// TwinCAT 3 PLC project PmsStd
// ProgramVersion: 3.1.4024.0
// libraries:
//   Tc3_IotBase, * (Beckhoff Automation GmbH)
//   Tc2_ModbusRTU, * (Beckhoff Automation GmbH)
//   Tc2_ModbusSrv, * (Beckhoff Automation GmbH)
//   Tc2_Standard, * (Beckhoff Automation GmbH)
//   Tc2_SUPS, * (Beckhoff Automation GmbH)
//   Tc2_System, * (Beckhoff Automation GmbH)
//   Tc3_Module, * (Beckhoff Automation GmbH)
//   Tc3_EventLogger, * (Beckhoff Automation GmbH)
//   Tc2_Utilities, * (Beckhoff Automation GmbH)
// project tree:
//   / FastTask.TcTTO, MqttTask.TcTTO, PlcTask.TcTTO, RedundancyTask.TcTTO
//   10_Core/00_Type/ ST_RuleTargetReg.TcDUT, ST_UnitLimitView.TcDUT, ST_BatLimitView.TcDUT, ST_BatLimitOut.TcDUT, ST_GateView.TcDUT, ST_GateOut.TcDUT, ST_SelectCand.TcDUT, ST_SelectView.TcDUT, ST_DistView.TcDUT, E_GridMode.TcDUT, ST_LogSet.TcDUT, E_StartMode.TcDUT, E_BatClose.TcDUT, ST_SeqSet.TcDUT, E_DistBasis.TcDUT, ST_CmdFilterSet.TcDUT, ST_RedSet.TcDUT, E_RedRole.TcDUT, ST_ModeSet.TcDUT, E_SelectMode.TcDUT, ST_GroupSet.TcDUT, ST_ManualPolicy.TcDUT, GVL_REASON.TcGVL, GVL_CORE.TcGVL, ST_UnitReq.TcDUT, ST_BmsCfg.TcDUT, E_PcsAction.TcDUT, E_BatAction.TcDUT, E_ModeAction.TcDUT, ST_ProtCfg.TcDUT, ST_PointTerm.TcDUT, ST_PointCfg.TcDUT, E_GroupState.TcDUT, E_LimitBasis.TcDUT, E_OpMode.TcDUT, E_ProtScope.TcDUT, E_RunState.TcDUT, E_SourceMode.TcDUT, ST_BatState.TcDUT, ST_GroupCfg.TcDUT, ST_GroupView.TcDUT, ST_Limit.TcDUT, ST_LimitOut.TcDUT, ST_MeterState.TcDUT, ST_ModuleReg.TcDUT, ST_PQ.TcDUT, ST_PccMeas.TcDUT, ST_RuleCfg.TcDUT, ST_SourceOutput.TcDUT, ST_SourceReg.TcDUT, E_PcsCmd.TcDUT, E_BatCmd.TcDUT, ST_PcsCmd.TcDUT, ST_BatCmd.TcDUT, ST_PcsReq.TcDUT, ST_BatReq.TcDUT, ST_PcsSeqSet.TcDUT, ST_BatSeqSet.TcDUT, ST_ManualCmdSet.TcDUT, ST_StateModeSet.TcDUT, ST_PcsCmdMode.TcDUT, ST_BatCmdMode.TcDUT, ST_UnitCfg.TcDUT, ST_UnitState.TcDUT, ST_Val.TcDUT, ST_OutputCfg.TcDUT, ST_ProtReq.TcDUT, ST_ProtView.TcDUT, E_CtrlModeRefuse.TcDUT, E_CtrlModeStep.TcDUT, ST_CtrlModeOut.TcDUT, ST_CtrlModeSet.TcDUT, ST_LocalTime.TcDUT, ST_CtrlModeView.TcDUT, E_PccShare.TcDUT, ST_UnitView.TcDUT
//   10_Core/01_Interface/ I_UnitLimitRule.TcIO, I_BatLimitRule.TcIO, I_Gate.TcIO, I_SelectPolicy.TcIO, I_DistPolicy.TcIO, I_AuxDevice.TcIO, I_OutputRule.TcIO, I_Bms.TcIO, I_CommandSource.TcIO, I_Compensator.TcIO, I_LimitRule.TcIO, I_Meter.TcIO, I_Module.TcIO, I_Pcs.TcIO, I_ReqDevice.TcIO, I_ProtResponse.TcIO, I_ProtectionRule.TcIO, I_StartPermit.TcIO, I_ControlMode.TcIO
//   10_Core/40_Arbitration/ FB_GateAuto.TcPOU, FB_GateManual.TcPOU, FB_SelectStd.TcPOU, F_RangeAnd.TcPOU, FB_PermitEval.TcPOU, FB_OutputReady.TcPOU, E_ModeSwitch.TcDUT, E_ModeStep.TcDUT, E_CmdRefuse.TcDUT, F_CmdOk.TcPOU, FB_ModeSwitch.TcPOU, FB_Gate.TcPOU, E_UnitRole.TcDUT, ST_Pick.TcDUT, ST_Range.TcDUT, ST_Clamp.TcDUT, ST_ShapeDiag.TcDUT, F_LimitKeepZero.TcPOU, F_RangeOpen.TcPOU, F_RangeAdd.TcPOU, F_RangeClamp.TcPOU, F_MakeLimit.TcPOU, F_SourceAllowed.TcPOU, F_StateRank.TcPOU, F_Better.TcPOU, FB_StateArbiter.TcPOU, FB_Select.TcPOU, FB_LimitEval.TcPOU, FB_ShapePath.TcPOU, F_PcsCmdAllowed.TcPOU, F_BatCmdAllowed.TcPOU
//   10_Core/50_Distribution/ FB_DistStd.TcPOU, E_UnitLimitBy.TcDUT, ST_UnitDiag.TcDUT, ST_DistDiag.TcDUT, ST_DistPathDiag.TcDUT, ST_BatDistDiag.TcDUT, FB_Distributor.TcPOU
//   10_Core/20_Protection/ ST_UnitEnvelope.TcDUT, ST_BatEnvelope.TcDUT, ST_GroupEnvelope.TcDUT, FB_EquipmentLimits.TcPOU, ST_BmsProt.TcDUT, ST_BmsAvail.TcDUT, ST_BatGroupState.TcDUT, FB_BatGroup.TcPOU, ST_UnitProt.TcDUT, ST_UnitAvail.TcDUT, F_PcsRank.TcPOU, F_BatRank.TcPOU, FB_Protection.TcPOU, FB_UnitAvail.TcPOU
//   20_Module/Common/ ST_SocLimitSet.TcDUT, ST_RuleBitSet.TcDUT, ST_RuleValueSet.TcDUT, FB_BreakerCtrl.TcPOU, ST_UnitLimitSet.TcDUT, ST_UnitLimitItem.TcDUT, FB_UnitLimit.TcPOU, ST_BreakerSet.TcDUT, F_SocDerate.TcPOU, FB_SocLimit.TcPOU, FB_AuxIo.TcPOU, FB_RuleBit.TcPOU, FB_RuleValue.TcPOU, F_SocLimitSetErr.TcPOU, FB_LocalClock.TcPOU, F_WordsToReal.TcPOU, ST_TempHumState.TcDUT
//   90_Project/ ST_ModuleSet.TcDUT, GVL_TEST.TcGVL, GVL_MQTT.TcGVL, GVL_PARAM.TcGVL, GVL_PERSIST.TcGVL, GVL_SITE.TcGVL, MAIN.TcPOU, GVL_IF.TcGVL, PRG_Mqtt.TcPOU, PRG_Fast.TcPOU, PRG_Redundancy.TcPOU
//   10_Core/60_Dispatch/ FB_GroupState.TcPOU, FB_BatRequest.TcPOU, E_UnitSeq.TcDUT, E_SeqRefuse.TcDUT, F_CmdReached.TcPOU, FB_UnitSeq.TcPOU, FB_BmsSeq.TcPOU, FB_Sequencer.TcPOU, FB_Dispatcher.TcPOU, FB_AuxOutput.TcPOU
//   10_Core/70_Diag/ FB_SettingGuard.TcPOU, FB_ModuleList.TcPOU, E_DiagStage.TcDUT, ST_OutputDiag.TcDUT, E_TraceStep.TcDUT, ST_TraceStep.TcDUT, ST_PTrace.TcDUT, F_TxtPcsAction.TcPOU, F_TxtBatAction.TcPOU, F_TxtSeq.TcPOU, F_TxtRefuse.TcPOU, F_TxtLimitBy.TcPOU, F_TxtStage.TcPOU, F_TxtOpMode.TcPOU, F_TxtCoreReason.TcPOU, F_TxtNum.TcPOU, FB_LogAlarm.TcPOU, FB_LogMsg.TcPOU, FB_OutputDiag.TcPOU, FB_AliveRecorder.TcPOU, FB_EventLog.TcPOU, FB_ConfigCheck.TcPOU, F_TxtPcsCmd.TcPOU, F_TxtBatCmd.TcPOU
//   10_Core/80_Report/ FB_Report.TcPOU
//   10_Core/02_Util/ F_ModeApplies.TcPOU, F_RampStep.TcPOU, FB_Lpf.TcPOU, FB_PersistSave.TcPOU, FB_ReadTimer.TcPOU, F_CycleSec.TcPOU, F_IsStopped.TcPOU, F_IsLocal.TcPOU, F_TimeHhmm.TcPOU, F_RealChanged.TcPOU, F_RealOk.TcPOU, F_RealToDint.TcPOU, F_HhmmOk.TcPOU, F_InHhmmWindow.TcPOU, F_MinutesTo.TcPOU, F_IsFinite.TcPOU
//   10_Core/30_Request/ FB_GroupView.TcPOU, FB_SourceHub.TcPOU, FB_CtrlModeMgr.TcPOU, FB_UnitView.TcPOU
//   20_Module/Standard/ FB_ProtRespStd.TcPOU, FB_ProtPcsFault.TcPOU, FB_ProtPcsComm.TcPOU, FB_ProtBmsFault.TcPOU, FB_ProtBmsComm.TcPOU, FB_ProtPccInvalid.TcPOU
//   10_Core/10_Snapshot/ ST_VirtualSet.TcDUT, FB_Snapshot.TcPOU, FB_Measure.TcPOU
//   10_Core/03_Base/ FB_DeviceBase.TcPOU, FB_ModuleBase.TcPOU, FB_SourceBase.TcPOU, FB_CtrlModeBase.TcPOU
//   20_Module/Mqtt/ FB_MqttPublish.TcPOU, FB_MqttSubscribe.TcPOU, F_MqttDistribute.TcPOU, PRG_PublishDeviceNo.TcPOU, ST_MqttCommand_Rx.TcDUT, ST_MqttCommandHeader.TcDUT, ST_MqttHeader.TcDUT, ST_MqttPubEntry.TcDUT, ST_MqttSubEntry.TcDUT, ST_IfEmsCmd.TcDUT, FB_EmsCommand.TcPOU, FB_SrcEms.TcPOU, FB_MqttMain.TcPOU, ST_MqttBroker.TcDUT, ST_MqttSet.TcDUT, ST_IfReport.TcDUT, F_MqttTimeText.TcPOU, FB_EmsConfigApply.TcPOU, FB_BrokerWatch.TcPOU, E_MqttBroker.TcDUT, ST_BrokerWatchSet.TcDUT, ST_IfEmsCfg.TcDUT, ST_IfEmsCfgEcho.TcDUT, ST_IfUpsConfigRx.TcDUT, FB_EmsCmdGate.TcPOU
//   20_Module/Mqtt/Publish/ ST_AirConditionerPublish_V1.TcDUT, ST_BatPublish_V1.TcDUT, ST_EssPublish_V1.TcDUT, ST_PcsPublish_V1.TcDUT, ST_PmsPublish_V1.TcDUT, ST_PvPublish_V1.TcDUT, ST_RackPublish_V1.TcDUT, ST_TempPublish_V1.TcDUT, ST_AirConditionerPublishData.TcDUT, ST_BatPublishData.TcDUT, ST_EssPublishData.TcDUT, ST_PcsPublishData.TcDUT, ST_PmsPublishData.TcDUT, ST_PvPublishData.TcDUT, ST_RackPublishData.TcDUT, ST_TempPublishData.TcDUT, ST_UpsPublish_V1.TcDUT, ST_ModulePublish_V1.TcDUT, ST_UpsPublishData.TcDUT, ST_ModulePublishData.TcDUT, ST_ImdPublish_V1.TcDUT, ST_ImdPublishData.TcDUT, ST_FirePublish_V1.TcDUT, ST_FirePublishData.TcDUT
//   20_Module/Mqtt/Config/ ST_BatConfig_Rx.TcDUT, ST_CommonConfig_REAL.TcDUT, ST_CommonConfig_UDINT.TcDUT, ST_PcsConfig_Rx.TcDUT, ST_ProtectionConfig_Rx.TcDUT, ST_BatConfigWirePacket.TcDUT, ST_PcsConfigWirePacket.TcDUT, ST_ProtectionConfigWirePacket.TcDUT, ST_UpsConfig_Rx.TcDUT, ST_UpsConfigWirePacket.TcDUT, ST_ScheduleWork_V1.TcDUT, ST_ScheduleHoliday_V1.TcDUT, ST_ScheduleDaily_V1.TcDUT, ST_ScheduleWeekly_V1.TcDUT
//   20_Module/Virtual/ PRG_MqttTestData.TcPOU, FB_BmsSim.TcPOU, FB_MeterSim.TcPOU, FB_PcsSim.TcPOU, FB_SrcTest.TcPOU, PRG_SimLink.TcPOU
//   20_Module/Mqtt/Logger/ FB_MqttLoggerListener.TcPOU, F_Utf8ToWstring.TcPOU, ST_LoggerHeader.TcDUT, ST_LoggerPublish_V1.TcDUT, ST_LoggerSlot.TcDUT
//   20_Module/Report/ FB_RptEsolutionBat.TcPOU, FB_RptSebangUps.TcPOU, FB_RptPlaspoPcs.TcPOU, FB_RptLsImd1000.TcPOU, FB_RptTempHum.TcPOU
//   20_Module/ControlMode/ ST_CmConstPowerSet.TcDUT, FB_CmConstPower.TcPOU, FB_CmStdSchedule.TcPOU, ST_CmExtCmd.TcDUT, ST_SchedSlot.TcDUT, ST_CmScheduleSet.TcDUT, FB_CmSchedule.TcPOU, GVL_CM_RSN.TcGVL, ST_CmDisWindow.TcDUT, ST_CmNoReverse.TcDUT, ST_CmCommonSet.TcDUT, ST_CmPeakCalcSet.TcDUT, ST_CmWindowSet.TcDUT, ST_CmPeakCutSet.TcDUT, ST_CmSchedPeakSet.TcDUT, F_CmVelocity.TcPOU, F_CmRoundTens.TcPOU, FB_CmTariffBase.TcPOU, FB_CmPeakCalc.TcPOU, FB_CmPeakCut.TcPOU, FB_CmSchedPeak.TcPOU
//   99_Test/ FB_TestTally.TcPOU, PRG_TestCtrlMode.TcPOU, PRG_TestSchedLive.TcPOU, PRG_TestPeakLive.TcPOU, PRG_TestUnitMode.TcPOU, PRG_TestStdLive.TcPOU, PRG_TestLogger.TcPOU, ST_LoggerTestReg.TcDUT
//   20_Module/Driver/Plaspo/ ST_PlaspoPcsRaw.TcDUT, FB_PlaspoPcs.TcPOU
//   10_Core/90_Redundancy/ E_RedPeer.TcDUT, ST_RedHeartbeat.TcDUT, FB_RedPeerMonitor.TcPOU, FB_RedLink.TcPOU, E_RedState.TcDUT, FB_RedState.TcPOU, E_RedSwitch.TcDUT, ST_RedSyncCfg.TcDUT, FB_RedSync.TcPOU
//   20_Module/Ups/ E_UpsResult.TcDUT, ST_UpsState.TcDUT, F_UpsSignedWord.TcPOU, F_UpsNextSeq.TcPOU, FB_UpsConfigApply.TcPOU, FB_UpsModbusJob.TcPOU, I_Ups.TcIO, E_UpsChargeAction.TcDUT, E_UpsChargeMode.TcDUT, E_UpsChargeStep.TcDUT, FB_UpsChargeRequest.TcPOU, FB_UpsChargeSequence.TcPOU, FB_UpsTemperatureCharge.TcPOU, ST_UpsChargeFeedback.TcDUT, ST_UpsChargeRequest.TcDUT, ST_UpsChargeSet.TcDUT, FB_UpsSafetyStage.TcPOU, ST_UpsDesiredSet.TcDUT, ST_IfUpsCmd.TcDUT, FB_UpsCommand.TcPOU, FB_UpsSafetyResponse.TcPOU, FB_UpsSafetyLog.TcPOU
//   20_Module/Driver/Sebang/ E_UpsCommand.TcDUT, ST_UpsRaw.TcDUT, F_DecodeSebangUps.TcPOU, FB_SebangUps.TcPOU
//   20_Module/Driver/Esolution/ E_EsolutionOperation.TcDUT, ST_EsolutionRaw.TcDUT, ST_EsolutionState.TcDUT, FB_EsolutionBms.TcPOU, E_EsolutionControl.TcDUT, ST_BatRackCmd.TcDUT, FB_BmsRackCommand.TcPOU, ST_BatCtlCmd.TcDUT, FB_BmsContactorCommand.TcPOU
//   20_Module/Driver/Autonics/ FB_AutonicsThd.TcPOU
//   20_Module/Driver/Bender/ FB_BenderIso685.TcPOU
//   20_Module/Driver/Rootech/ FB_RootechAcuraIo.TcPOU
//   20_Module/Driver/LS/ ST_LsImd1000State.TcDUT, FB_LsImd1000.TcPOU
//   20_Module/Driver/ITGuard/ FB_ItGuardIeSx.TcPOU
//   20_Module/Driver/Woonyoung/ FB_WoonyoungGfr.TcPOU
//   20_Module/Driver/Gasdna/ FB_GasdnaAsd57.TcPOU
// real-time tasks:
//   TASK PlcTask: cycle T#10ms, priority 20, ADS port 350
//   TASK MqttTask: cycle T#10ms, priority 30, ADS port 351
//   TASK FastTask: cycle T#10ms, priority 2, ADS port 352
//   TASK RedundancyTask: cycle T#10ms, priority 1, ADS port 353
// I/O:
//   DEVICE Device 1 (EtherCAT Automation Protocol), AmsNetId 10.1.177.153.2.1
//     Box 2 (Subscriber)
//     Box 1 (Publisher)
//   DEVICE Device 2 (EtherCAT), AmsNetId 10.1.177.153.3.1
//     Term 1 (EK1200) [EK1200-5000 EtherCAT Power supply (2A E-Bus)]
//       Term 4 (EL1004) [EL1004 4Ch. Dig. Input 24V, 3ms]
//       Term 5 (EL2004) [EL2004 4Ch. Dig. Output 24V, 0.5A]
//       Term 6 (EL6022) [EL6022 Interface 2Ch. (RS422/485)]
//       Term 5 (EL9011) [EL9011 End Terminal]
// variable links:
//   PmsStd/PmsStd Instance <-> Device 1 (EtherCAT Automation Protocol)/Box 1 (Publisher)
//     RedundancyTask Outputs/PRG_Redundancy.fbRedLink._stTx <-> RedHeartbeat/Outputs/VarData
//     RedundancyTask Outputs/PRG_Redundancy.fbRedSync._stTx <-> RedSyncCfg/Outputs/VarData
//   PmsStd/PmsStd Instance <-> Device 1 (EtherCAT Automation Protocol)/Box 2 (Subscriber)
//     RedundancyTask Inputs/PRG_Redundancy.fbRedLink._nEapQuality <-> RedHeartbeat/Inputs/Quality
//     RedundancyTask Inputs/PRG_Redundancy.fbRedLink._stRx <-> RedHeartbeat/Inputs/VarData
//     RedundancyTask Inputs/PRG_Redundancy.fbRedSync._stRx <-> RedSyncCfg/Inputs/VarData
//   PmsStd/PmsStd Instance <-> Device 2 (EtherCAT)/Term 1 (EK1200)/Term 4 (EL1004)
//     RedundancyTask Inputs/PRG_Redundancy.fbRedLink._bDiPeerActive <-> Channel 2/Input
//     RedundancyTask Inputs/PRG_Redundancy.fbRedLink._bDiPeerAlive <-> Channel 1/Input
//   PmsStd/PmsStd Instance <-> Device 2 (EtherCAT)/Term 1 (EK1200)/Term 5 (EL2004)
//     RedundancyTask Outputs/PRG_Redundancy.fbRedLink._bDoActive <-> Channel 2/Output
//     RedundancyTask Outputs/PRG_Redundancy.fbRedLink._bDoAlive <-> Channel 1/Output

CONFIGURATION PmsStd
    RESOURCE PLC ON TwinCAT3
        TASK FastTask(INTERVAL := T#10ms, PRIORITY := 2);
        TASK MqttTask(INTERVAL := T#10ms, PRIORITY := 30);
        TASK PlcTask(INTERVAL := T#10ms, PRIORITY := 20);
        TASK RedundancyTask(INTERVAL := T#10ms, PRIORITY := 1);
        PROGRAM PRG_Fast WITH FastTask : PRG_Fast;
        PROGRAM PRG_Mqtt WITH MqttTask : PRG_Mqtt;
        PROGRAM MAIN WITH PlcTask : MAIN;
        PROGRAM PRG_Redundancy WITH RedundancyTask : PRG_Redundancy;
    END_RESOURCE
END_CONFIGURATION

// ---- 10_Core/00_Type/ST_RuleTargetReg.TcDUT
TYPE ST_RuleTargetReg :	// 유닛 제한·버스 제한 모듈 등록 (칸 번호는 GVL_SITE 등록 배열과 같음)
STRUCT
	bEnable	: BOOL := TRUE;
	nTarget	: UINT;	// 대상 번호 (유닛 제한 = 유닛, 버스 제한 = 배터리 그룹). 0 = 전체 (모듈이 대상별 상태를 따로 가짐)
	bAuto	: BOOL := TRUE;	// Auto 유닛에 적용
	bManual	: BOOL := TRUE;	// Manual 유닛에 적용. 버스 제한은 그 버스에 적용 대상 모드 유닛이 하나라도 있으면 버스 전체에 걸림 (버스에 유닛이 없으면 그대로 걸림)
END_STRUCT
END_TYPE

// ---- 10_Core/00_Type/ST_UnitLimitView.TcDUT
TYPE ST_UnitLimitView :	// 유닛 제한 모듈에 넘기는 유닛 요약 (읽기 전용)
STRUCT
	nUnit	: UINT;
	eOpMode	: E_OpMode;	// 실제 운전 모드
	bAvail	: BOOL;
	eRunState	: E_RunState;
	stP	: ST_Val;	// kW, 실측
	stQ	: ST_Val;	// kvar, 실측
	fPRated	: REAL;	// kW
	fQRated	: REAL;	// kvar
	nBatGroup	: UINT;	// 연결 배터리 그룹. 0 = 없음
	stSoc	: ST_Val;	// %, 연결 배터리 그룹 평균
END_STRUCT
END_TYPE

// ---- 10_Core/00_Type/ST_BatLimitView.TcDUT
TYPE ST_BatLimitView :	// 버스 제한 모듈에 넘기는 배터리 그룹(DC 버스) 요약 (읽기 전용)
STRUCT
	nBatGroup	: UINT;
	bUsable	: BOOL;	// 쓸 수 있는 BMS가 하나 이상
	stSoc	: ST_Val;	// %, 용량 가중 평균
	stSocMin	: ST_Val;	// %
	stSocMax	: ST_Val;	// %
	fPChgMax	: REAL;	// kW, BMS 충전 한도 합 (양수)
	fPDisMax	: REAL;	// kW, BMS 방전 한도 합 (양수)
	fPOut	: REAL;	// kW, 이 버스 유닛 출력 합 (실측)
	nUnitAuto	: UINT;	// 이 버스의 Auto 유닛 수
	nUnitManual	: UINT;	// 이 버스의 Manual 유닛 수
END_STRUCT
END_TYPE

// ---- 10_Core/00_Type/ST_BatLimitOut.TcDUT
TYPE ST_BatLimitOut :	// 버스 제한 모듈 결과
STRUCT
	stP	: ST_Limit;	// kW. fMax = 방전 상한(0 이상), fMin = 충전 하한(0 이하). bActive = FALSE면 제한 없음
	bResume	: BOOL;	// 출력 재개 중: 코어 램프가 재개 램프율을 씀
END_STRUCT
END_TYPE

// ---- 10_Core/00_Type/ST_GateView.TcDUT
TYPE ST_GateView :	// Gate에 넘기는 것 (I_Gate.M_Filter)
STRUCT
	ePath			: E_OpMode;			// 이 Gate가 맡은 경로 (Auto / Manual)
	stManualCmdSet	: ST_ManualCmdSet;	// Manual 지령 거르기 설정 (GVL_PERSIST.g_stManualCmdSet, 코어 기본 Manual Gate가 씀)
END_STRUCT
END_TYPE

// ---- 10_Core/00_Type/ST_GateOut.TcDUT
TYPE ST_GateOut :	// Gate 결과: 성형·분배는 지령 값을, 디스패처·로그는 새 지령·거부·대기를 씀
STRUCT
	astUnitP		: ARRAY[1..GVL_PARAM.UNIT_COUNT] OF ST_Pick;		// 거른 유닛별 값
	astUnitQ		: ARRAY[1..GVL_PARAM.UNIT_COUNT] OF ST_Pick;
	astGrpP			: ARRAY[1..GVL_PARAM.GROUP_COUNT] OF ST_Pick;		// 거른 그룹 값
	astGrpQ			: ARRAY[1..GVL_PARAM.GROUP_COUNT] OF ST_Pick;
	abNew			: ARRAY[1..GVL_PARAM.UNIT_COUNT] OF BOOL;		// 새 지령을 받아들임 (Manual: 디스패처가 이 스캔에 바로 씀)
	aeRefuse		: ARRAY[1..GVL_PARAM.UNIT_COUNT] OF E_CmdRefuse;	// 마지막으로 무시한 이유 (받아들이면 None)
	anRefuseModule	: ARRAY[1..GVL_PARAM.UNIT_COUNT] OF UINT;		// 무시한 지령을 낸 모듈 ID
	abWaitNewCmd	: ARRAY[1..GVL_PARAM.UNIT_COUNT] OF BOOL;		// 새 지령이 올 때까지 출력 0 (Manual)
END_STRUCT
END_TYPE

// ---- 10_Core/00_Type/ST_SelectCand.TcDUT
TYPE ST_SelectCand :	// 고르기 후보 하나 (지령원 하나의 값)
STRUCT
	nSource		: UINT;		// 지령원 칸 번호 (g_aipSource)
	nModule		: UINT;		// 지령원 모듈 ID
	nGrade		: UINT;		// 등급 (1이 가장 높음, g_astSourceReg)
	fValue		: REAL;		// kW 또는 kvar (이상값은 코어가 미리 뺌)
	bNew		: BOOL;		// 이번 스캔에 새 지령
END_STRUCT
END_TYPE

// ---- 10_Core/00_Type/ST_SelectView.TcDUT
TYPE ST_SelectView :	// 고르기 정책에 넘기는 것 (I_SelectPolicy.M_Select). 후보는 지령원 칸 순서
STRUCT
	nGroup		: UINT;			// 제어 그룹
	nUnit		: UINT;			// 0 = 그룹 값, n = 유닛 n의 유닛별 값
	bForQ		: BOOL;			// FALSE = P, TRUE = Q
	eOpMode		: E_OpMode;		// 경로 (Auto / Manual). 유닛별 값이면 그 유닛의 운전 모드
	eSel		: E_SelectMode;	// 그룹 설정 eSelP·eSelQ (기본 정책이 씀)
	nCand		: UINT;			// 후보 수
	astCand		: ARRAY[1..GVL_PARAM.SOURCE_COUNT] OF ST_SelectCand;	// 1..nCand만 유효
END_STRUCT
END_TYPE

// ---- 10_Core/00_Type/ST_DistView.TcDUT
TYPE ST_DistView :	// 분배 정책에 넘기는 것 (I_DistPolicy.M_Weight): 유닛 하나
STRUCT
	nGroup		: UINT;
	nUnit		: UINT;
	bManual		: BOOL;			// Manual 경로 그룹 몫
	bForQ		: BOOL;			// FALSE = P, TRUE = Q
	bPositive	: BOOL;			// 나눌 양이 방전·공급 쪽
	eBasis		: E_DistBasis;	// 그룹 설정 eDistBasis (기본 정책이 씀)
	fPRated		: REAL;			// kW, 정격 (Derate 반영 전)
	fQRated		: REAL;			// kvar
	fSoc		: REAL;			// %, 연결 배터리 그룹 SOC. 모르면 -1
END_STRUCT
END_TYPE

// ---- 10_Core/20_Protection/ST_UnitEnvelope.TcDUT
TYPE ST_UnitEnvelope :	// 유닛 설비 한도 (FB_EquipmentLimits). 가용·운전 상태와 관계없는 장비 한도
STRUCT
	stP	: ST_Range;	// kW. 정격 × Derate ∩ 유닛 제한 모듈 (모듈 0 = 코어). 0은 항상 범위 안
	stQ	: ST_Range;	// kvar
	stPRule	: ST_Range;	// kW. 유닛 제한 모듈만 (Manual 정책 bRating을 끈 유닛에 씀)
	stQRule	: ST_Range;	// kvar
	fSMax	: REAL;	// kVA, 피상전력 한도 = MIN(정격 S, √(보호 P 상한² + 보호 Q 상한²))
	bDerated	: BOOL;	// 보호 Derate 걸림
	ePMaxBy	: E_UnitLimitBy;	// P 상한을 정한 것: Rating / Derate / UnitRule
	ePMinBy	: E_UnitLimitBy;	// P 하한을 정한 것
	eQMaxBy	: E_UnitLimitBy;
	eQMinBy	: E_UnitLimitBy;
	bResume	: BOOL;	// 유닛 제한 모듈이 재개 중
END_STRUCT
END_TYPE

// ---- 10_Core/20_Protection/ST_BatEnvelope.TcDUT
TYPE ST_BatEnvelope :	// 배터리 그룹(DC 버스) 한도 (FB_EquipmentLimits)
STRUCT
	stP	: ST_Range;	// kW. fMax = 방전 한도(0 이상), fMin = -충전 한도(0 이하). BMS 한도 합 ∩ 버스 제한 모듈 (모듈 0 = BMS 한도)
	bResume	: BOOL;	// 버스 제한 모듈이 재개 중
END_STRUCT
END_TYPE

// ---- 10_Core/20_Protection/ST_GroupEnvelope.TcDUT
TYPE ST_GroupEnvelope :	// 제어 그룹 설비 범위 (가용 유닛 기준). 성형의 설비 제한 줄 (정격·배터리)
STRUCT
	stRating	: ST_Range;	// kW, 가용 유닛 P 한도 합 (정격 × Derate ∩ 유닛 제한 모듈)
	stBattery	: ST_Range;	// kW, 버스마다 min(버스 한도, 그 버스 가용 유닛 한도 합) + 배터리 없는 유닛 한도
	stQ	: ST_Range;	// kvar, 가용 유닛 Q 한도 합
	fSMax	: REAL;	// kVA, 가용 유닛 피상전력 한도 합 (유닛 한도 = MIN(정격 S, √(보호 P 상한² + 보호 Q 상한²)))
	bResume	: BOOL;	// 유닛·버스 제한 모듈이 재개 중 (재개 램프율)
END_STRUCT
END_TYPE

// ---- 20_Module/Common/ST_SocLimitSet.TcDUT
TYPE ST_SocLimitSet :	// FB_SocLimit 설정 (운전 중 HMI로 바꿈. GVL_PERSIST.g_stModuleSet 칸 → MAIN이 매 스캔 넘김)
STRUCT
	fSocMax	: REAL := 95.0;	// %, 이 값 이상이면 충전 막음
	fSocMin	: REAL := 5.0;	// %, 이 값 이하면 방전 막음
	fBand	: REAL := 5.0;	// %, 한계 앞 이 폭에서 한도를 선형으로 줄임. 0 = 줄이지 않고 한계에서 막기만
	fResumeMargin	: REAL := 2.0;	// %, 막은 뒤 한계에서 이만큼 돌아와야 다시 허용 (재개 마진)
	bBlockOnInvalid	: BOOL := TRUE;	// SOC 무효면 충·방전 모두 막음
END_STRUCT
END_TYPE

// ---- 20_Module/Common/ST_RuleBitSet.TcDUT
TYPE ST_RuleBitSet :	// FB_RuleBit 설정 (운전 중 HMI로 바꿈. GVL_PERSIST.g_stModuleSet 칸 → MAIN이 매 스캔 넘김)
STRUCT
	bInvert	: BOOL;	// TRUE = b접점 (평소 닫힘, 열리면 조건)
	bOnCommLoss	: BOOL;	// 보조 장비 통신(I/O)이 끊기면 조건 있음으로 봄
END_STRUCT
END_TYPE

// ---- 20_Module/Common/ST_RuleValueSet.TcDUT
TYPE ST_RuleValueSet :	// FB_RuleValue 설정 (운전 중 HMI로 바꿈. 임계값은 등록 설정 fThreshold. GVL_PERSIST.g_stModuleSet 칸 → MAIN이 매 스캔 넘김)
STRUCT
	bBelow	: BOOL;	// FALSE = 임계값 이상이면 조건, TRUE = 이하면 조건
	fHyst	: REAL;	// 해소 폭: 임계값에서 이만큼 돌아와야 풀림
	bOnCommLoss	: BOOL;	// 통신이 끊기거나 값이 무효면 조건 있음으로 봄
END_STRUCT
END_TYPE

// ---- 90_Project/ST_ModuleSet.TcDUT
TYPE ST_ModuleSet :	// 현장 모듈 설정 묶음 (GVL_PERSIST.g_stModuleSet). 운전 중 HMI로 바꾸고 재기동해도 유지
// 현장에 모듈을 추가하면: 여기 칸 추가 → MAIN 액션 A_PassModuleSet에 한 줄 추가 (저장·잘못된 값 되돌리기는 묶음 전체를 봄)
STRUCT
	stSocLimit	: ST_SocLimitSet;	// g_fbSocLimit: 기본 SOC 95 / 5 %, 감발 폭 5 %, 재개 마진 2 %, SOC 무효면 막음
	(* 제어 모드: 접속점 그룹 1 관리자(g_fbCtrlMode1, 접속점 그룹 단위)와 모드 한 세트. 공통(월 → 계절, 휴일, 방전 허용 시간 월~토 08~22시, 역송 방지 여유 10 kW)은 stCmCommon
	   [16번 수정 2026-11-09: PCS2 칸(stCtrlMode2·stCmConstP2·stCmSchedule2·stCmPeakCut2·stCmSchedPeak2) 없앰. 값은 접속점 그룹 전체 기준 (피크 목표·정출력 = 접속점 그룹의 접속점 값)] *)
	stCmCommon		: ST_CmCommonSet;
	stCtrlMode1		: ST_CtrlModeSet := (bZeroOnSwitch := TRUE, tZeroDelay := T#1S, nFallback := 0, ePccShare := E_PccShare.ByRating, fPccRatio := 1.0);	// g_fbCtrlMode1: 바꿀 때 1 s 출력 0, 스스로 끝나면 모드 없음 (ePccShare·fPccRatio는 유닛 단위 관리자만 씀)
	stCmConstP1		: ST_CmConstPowerSet := (fPSet := 0.0, bQSet := FALSE, fQSet := 0.0, tDuration := T#0S);	// g_fbCmConstP1: fPSet (kW, 방전 +, 접속점 그룹의 접속점 기준)
	stCmSchedule1	: ST_CmScheduleSet;		// 접속점 그룹 1 시간표 [계절, 요일, 칸] (kW, 방전 +, 접속점 그룹 값). 스케줄·통합이 같이 씀. 기본 = 빈 시간표 (0을 냄)
	stCmPeakCut1		: ST_CmPeakCutSet;		// g_fbCmPeakCut1: 목표 피크 stPeak.fTarget (kW, 접속점 그룹 전체. 0 = 제어 안 함), 자동 충전·잔량 방전 시간 (기본 끔)
	stCmSchedPeak1	: ST_CmSchedPeakSet;	// g_fbCmSchedPeak1: 목표 피크 (접속점 그룹 전체), 잔량 방전 시간 (기본 끔)
	stUnitLimit	: ST_UnitLimitSet;	// g_fbUnitLimit 사용자 한도 (유닛마다 P·Q 상·하한 kW·kvar). 기본: 모두 끔. HMI 또는 EMS config pcs(FB_EmsConfigApply)가 씀 [9-21 수정 2026-11-04: 아래 주석 예에서 꺼냄 (맨 끝에 붙여 앞 칸 배치는 그대로)]
	(* 예 (GVL_SITE 주석 예와 같이 풀어 씀)
	stFire	: ST_RuleBitSet;
	stEStop	: ST_RuleBitSet := (bInvert := TRUE, bOnCommLoss := TRUE);
	stBatTemp	: ST_RuleValueSet := (fHyst := 2.0);
	stVcb1	: ST_BreakerSet := (tPulse := T#1S, tConfirm := T#5S);
	(9-21 수정 2026-11-04: stUnitLimit은 위로 꺼냄) stUnitLimit	: ST_UnitLimitSet;	// 기본: 모두 끔. HMI에서 astUnit[n].bPEnable·fPMax·fPMin (kW) 등을 바꿈
	*)
END_STRUCT
END_TYPE

// ---- 10_Core/00_Type/E_GridMode.TcDUT
{attribute 'qualified_only'}
{attribute 'strict'}
TYPE E_GridMode :		// PCS 계통 제어 방식 (유닛 속성. Auto/Manual처럼 경로를 가르지 않음)
(
	Unknown		:= 0,	// 모름
	Gfl			:= 1,	// 계통 추종 (Grid Following, 기본)
	Gfm			:= 2	// 계통 형성 (Grid Forming). 계통 연계 중에는 PMS 계산이 같음 (P·Q 지령, 전압·주파수 드룹은 PCS가 처리)
) INT;
END_TYPE

// ---- 20_Module/Common/ST_UnitLimitSet.TcDUT
TYPE ST_UnitLimitSet :	// FB_UnitLimit 설정 (운전 중 HMI로 바꿈. GVL_PERSIST.g_stModuleSet 칸 → MAIN A_PassModuleSet이 넘김)
STRUCT
	astUnit		: ARRAY[1..GVL_PARAM.UNIT_COUNT] OF ST_UnitLimitItem;	// 유닛마다 (기본: 모두 끔)
END_STRUCT
END_TYPE

// ---- 20_Module/Common/ST_UnitLimitItem.TcDUT
TYPE ST_UnitLimitItem :	// 유닛 하나의 사용자 한도 (kW·kvar)
STRUCT
	bPEnable	: BOOL;			// P 한도 사용
	fPMax		: REAL;			// kW, 방전 상한 (0 이상)
	fPMin		: REAL;			// kW, 충전 하한 (0 이하. 예: -500 = 충전 500 kW까지)
	bQEnable	: BOOL;			// Q 한도 사용
	fQMax		: REAL;			// kvar, 공급 상한 (0 이상)
	fQMin		: REAL;			// kvar, 흡수 하한 (0 이하)
END_STRUCT
END_TYPE

// ---- 20_Module/Common/ST_BreakerSet.TcDUT
TYPE ST_BreakerSet :	// FB_BreakerCtrl 설정 (운전 중 HMI로 바꿈. GVL_PERSIST.g_stModuleSet 칸 → MAIN A_PassModuleSet이 넘김)
STRUCT
	tPulse		: TIME := T#1S;		// 코일 펄스 폭 (투입·개방)
	tConfirm	: TIME := T#5S;		// 지령 뒤 이 시간 안에 상태 접점이 바뀌어야 함 (아니면 실패)
END_STRUCT
END_TYPE

// ---- 10_Core/00_Type/ST_LogSet.TcDUT
TYPE ST_LogSet :
STRUCT
	tHold			: TIME := T#10S;	// 출력 제한 이유가 이 시간 이상 유지될 때만 기록
	tPersistSave	: TIME := T#60S;	// PERSISTENT 주기 저장 (재기동 기록 시각 포함. 설정 변경은 바로 저장)
	bCmdRefused		: BOOL := TRUE;		// 무시한 지령 기록 (이상값·방향 반대·운전 모드 설정·보호 중 버린 요청)
	bBatRefused		: BOOL := TRUE;		// 배터리 요청 거부 (잠금·버스 유닛 운전 중) 기록
	(* 자세한 기록: 기본 끔 (시운전·문제 추적 때 켬) *)
	bUnitLimited	: BOOL;
	bReqRefused		: BOOL;
	bSeqChange		: BOOL;
	bModeChange		: BOOL;
END_STRUCT
END_TYPE

// ---- 10_Core/70_Diag/E_DiagStage.TcDUT
{attribute 'qualified_only'}
{attribute 'strict'}
TYPE E_DiagStage :
(
	None		:= 0,	// 요청대로 나감
	NoRequest	:= 1,	// 출력 요청 없음 (정상)
	NotRunning	:= 2,	// 그룹이 운전 중 아님
	Ramp		:= 3,	// 램프로 따라가는 중
	PccLimit	:= 4,	// 접속점 제한
	DeviceLimit	:= 5,	// 설비 제한 (정격·배터리·설비 기준 모듈)
	UnitLimit	:= 6,	// 유닛 한도·분배
	NoUnit		:= 7	// 그룹에 이 모드(Auto/Manual) 유닛이 없음 (정상, 로그 안 남김)
) INT;
END_TYPE

// ---- 10_Core/70_Diag/ST_OutputDiag.TcDUT
TYPE ST_OutputDiag :
STRUCT
	eStage		: E_DiagStage;		// 막은 단계. Auto P: 최종 값을 정한 단계 (추적표 기준), 나머지: 처음 막은 단계
	nModule		: UINT;				// 막은 모듈 (0 = 코어)
	nReason		: UINT;				// 이유 코드 (모듈이 정한 이유 또는 GVL_REASON 코어 이유). UnitLimit 단계는 0
	eUnitBy		: E_UnitLimitBy;	// UnitLimit 단계일 때 유닛 한도 이유 (그 경로 유닛 중 처음 찾은 것)
	eGroupState	: E_GroupState;		// NotRunning일 때 그룹 상태
	fReq		: REAL;				// kW, 고른 요청값
	fOut		: REAL;				// kW, 장비에 쓴 값 합
END_STRUCT
END_TYPE

// ---- 10_Core/70_Diag/E_TraceStep.TcDUT
{attribute 'qualified_only'}
{attribute 'strict'}
TYPE E_TraceStep :
(
	None		:= 0,
	Request		:= 1,	// 요청: 그룹 지령 또는 유닛 지령 합 (접속점 기준)
	Ramp		:= 2,	// 램프 후
	PccLimit	:= 3,	// 접속점 제한: 지령원 P 제한 또는 접속점 기준 모듈 하나
	Comp		:= 4,	// 보정을 더한 값 (여기부터 설비 기준)
	DevRating	:= 5,	// 설비 제한: 가용 정격
	DevBattery	:= 6,	// 설비 제한: 배터리 충·방전 한도
	DevLimit	:= 7,	// 설비 제한: 설비 기준 모듈 하나
	UnitDist	:= 8,	// 유닛 한도·분배 후 그룹 유닛 합
	Written		:= 9	// 장비에 쓴 값 합
) INT;
END_TYPE

// ---- 10_Core/70_Diag/ST_TraceStep.TcDUT
TYPE ST_TraceStep :		// 출력 추적표 한 줄
STRUCT
	eStep		: E_TraceStep;
	fValue		: REAL;			// kW, 이 단계를 지난 값
	bCut		: BOOL;			// 이 단계에서 값이 바뀜
	nModule		: UINT;			// 바꾼 모듈 (0 = 코어). Request 줄은 지령원 모듈
	nReason		: UINT;			// 이유 코드
END_STRUCT
END_TYPE

// ---- 10_Core/70_Diag/ST_PTrace.TcDUT
TYPE ST_PTrace :		// 출력 추적표 (P, 경로 하나·그룹 하나): 위에서부터 차례로 값이 어떻게 바뀌었는지
STRUCT
	nCount		: UINT;			// 채운 줄 수
	astStep		: ARRAY[1..GVL_PARAM.TRACE_STEP_MAX] OF ST_TraceStep;
END_STRUCT
END_TYPE

// ---- 10_Core/00_Type/E_StartMode.TcDUT
{attribute 'qualified_only'}
{attribute 'strict'}
TYPE E_StartMode :
(
	Step		:= 0,	// 단계별 기동: 작업자가 BatClose → Standby → Run을 하나씩 (기본, 지금 운영 방식)
	Sequence	:= 1	// 순서 기동: Run 요청 하나로 배터리 투입 → Standby → 기동 조건 → Run (운전 모드 Auto/Manual과 별개)
) INT;
END_TYPE

// ---- 10_Core/00_Type/E_BatClose.TcDUT
{attribute 'qualified_only'}
{attribute 'strict'}
TYPE E_BatClose :
(
	OnStart		:= 0,	// 순서 기동(E_StartMode.Sequence)하는 유닛이 있을 때 투입 (기본)
	OnRequest	:= 2	// 지령원의 BatClose 요청으로만 투입 (운전 모드 Manual과 별개)
) INT;
END_TYPE

// ---- 10_Core/00_Type/ST_SeqSet.TcDUT
TYPE ST_SeqSet :
STRUCT
	tWritePeriod	: TIME := T#200MS;		// Auto 유닛 P·Q 쓰기 주기 (Manual 유닛의 램프·설비 제한 추종도 이 주기)
	stPcs			: ST_PcsSeqSet;			// PCS(유닛) 시퀀스
	stBat			: ST_BatSeqSet;			// 배터리 시퀀스
END_STRUCT
END_TYPE

// ---- 10_Core/60_Dispatch/E_UnitSeq.TcDUT
{attribute 'qualified_only'}
{attribute 'strict'}
TYPE E_UnitSeq :
(
	Unknown		:= 0,	// 통신 전
	Stopped		:= 1,
	WaitBat		:= 2,	// 배터리 투입 대기 (순서 기동)
	Standby		:= 4,	// 대기 (활성 + 출력 0)
	WaitPermit	:= 5,	// 기동 조건 대기
	ToRun		:= 6,	// Run 명령 확인 중
	Running		:= 7,
	StopRamp	:= 8,	// 정지 전 출력 내리는 중
	ToStop		:= 9	// 정지 쪽 명령 보낼 차례(통신 대기)·확인 중
) INT;
END_TYPE

// ---- 10_Core/60_Dispatch/E_SeqRefuse.TcDUT
{attribute 'qualified_only'}
{attribute 'strict'}
TYPE E_SeqRefuse :
(
	None		:= 0,
	NotAvail	:= 1,	// 유닛이 가용 아님 (고장·통신·보호 등)
	NoBattery	:= 2,	// 배터리 미투입
	NoPermit	:= 4,	// 기동 조건 미충족
	CommLost	:= 6,	// 통신 없음
	UnitRunning	:= 8,	// 배터리 개방 요청인데 버스의 유닛이 정지 안 됨
	StopInProgress	:= 9,	// 정지 쪽 명령(Standby·Stop·EStop) 진행 중: 끝날 때까지 기동 요청 안 받음
	ConfigError	:= 10,	// 설정 오류로 장비 제어 중지 중
	WriteDisabled	:= 11	// 장비 쓰기 불가 (GVL_SITE.DEVICE_WRITE 꺼짐 또는 대기 PLC)
) INT;
END_TYPE

// ---- 10_Core/00_Type/E_DistBasis.TcDUT
{attribute 'qualified_only'}
{attribute 'strict'}
TYPE E_DistBasis :
(
	Rating		:= 0,	// 유닛 정격 비율
	Soc			:= 1,	// 방전은 SOC 높은 쪽, 충전은 SOC 낮은 쪽이 많이 (P만. Q는 정격 비율)
	Equal		:= 2	// 균등
) INT;
END_TYPE

// ---- 10_Core/50_Distribution/E_UnitLimitBy.TcDUT
{attribute 'qualified_only'}
{attribute 'strict'}
TYPE E_UnitLimitBy :
(
	None		:= 0,
	NotAvail	:= 1,	// 가용 아님 → 0
	NotRun		:= 2,	// 장비가 활성(Run·대기)이 아니거나 정지 진행 중 → 0
	Rating		:= 3,	// 유닛 정격
	Derate		:= 4,	// 보호 Derate
	Scaled		:= 5,	// 유닛별 값을 그룹 목표에 맞춰 비율로 줄임
	BatDir		:= 6,	// 같은 배터리 그룹의 순 방향과 반대 → 0
	BatLimit	:= 7,	// 배터리 버스 한도 (그 방향 한도 0, 버스 제한 모듈 포함)
	SLimit		:= 8,	// 피상전력 정격
	ModeSwitch	:= 9,	// 운전 모드 전환 중 → 0
	WaitManualCmd	:= 10,	// Manual: Run에서 빠졌다 돌아옴 → 새 지령이 올 때까지 0
	UnitRule	:= 11	// 유닛 제한 모듈 (I_UnitLimitRule)
) INT;
END_TYPE

// ---- 10_Core/00_Type/ST_CmdFilterSet.TcDUT
TYPE ST_CmdFilterSet :		// 명령 필터 설정 (FB_Select, Auto·Manual 공통). Manual 전용은 ST_ManualCmdSet
STRUCT
	(* 이상값: NaN·무한대는 항상 무시. 켜면 정격 × 배수를 넘는 값도 무시 (Auto·Manual) *)
	bBadValue		: BOOL := TRUE;
	fBadFactor		: REAL := 1.5;			// 그룹 값은 그룹 유닛 정격 합, 유닛별 값은 유닛 정격 기준
END_STRUCT
END_TYPE

// ---- 10_Core/00_Type/ST_RedSet.TcDUT
TYPE ST_RedSet :		// 이중화 설정 (GVL_SITE.RED_SET). 두 PLC에 같은 프로그램을 넣고, 역할은 이 PLC의 AMS Net ID로 정함
STRUCT
	bUse			: BOOL;			// FALSE(기본) = 이중화 안 씀: 이 PLC가 Primary이고 항상 장비에 씀
	sPrimaryNetId	: T_AmsNetId;	// Primary PLC의 AMS Net ID (예 '5.69.107.242.1.1')
	sSecondaryNetId	: T_AmsNetId;	// Secondary PLC의 AMS Net ID
	tEapTimeout		: TIME := T#500MS;	// EAP 하트비트 카운터가 안 바뀌거나 Quality(갱신 안 된 시간)가 이 시간을 넘으면 EAP 끊김 (FB_RedPeerMonitor)
	tWireTimeout	: TIME := T#500MS;	// 상대 접점(alive) 신호가 이 시간 안 바뀌면 접점 끊김
	tTakeoverDelay	: TIME := T#500MS;	// 절체 안전 지연: 상대가 Lost로 판정된 뒤 Secondary가 이 시간 더 기다렸다가 Active가 됨
	tFailbackStable	: TIME := T#10S;	// 복귀 조건: 상대(Secondary)와 통신이 이 시간 동안 계속 정상이어야 Primary가 Active를 넘겨받기 시작
	tHandoverTimeout: TIME := T#3S;		// 넘겨받기를 시작한 뒤 이 시간 안에 상대가 Active를 내려놓지 않으면 포기하고 Standby로 돌아감
	tWriteHold		: TIME := T#1S;		// Active가 된 뒤 이 시간이 지나야 장비에 씀 (승격 직후 값이 안정되기를 기다림)
	tStartGrace		: TIME := T#3S;		// 시작 직후 이 시간 안에는 상대 신호를 못 봐도 Unknown (끊김으로 보지 않음)
END_STRUCT
END_TYPE

// ---- 10_Core/00_Type/E_RedRole.TcDUT
{attribute 'qualified_only'}
{attribute 'strict'}
TYPE E_RedRole :		// 이중화에서 이 PLC의 역할 (고정 신분. 지금 장비에 쓰는지는 GVL_IF.g_bRedActive)
(
	Reading		:= 0,	// 이 PLC Net ID를 읽는 중 (시작 직후)
	Primary		:= 1,	// 주로 쓰는 PLC. 이중화를 안 쓰면 항상 Primary
	Secondary	:= 2,	// 예비 PLC
	NoMatch		:= 3	// 이 PLC Net ID가 GVL_SITE.RED_SET의 Primary·Secondary 어느 쪽과도 다름 → 설정 오류
) INT;
END_TYPE

// ---- 10_Core/00_Type/ST_ModeSet.TcDUT
TYPE ST_ModeSet :		// 운전 모드 전환 설정
STRUCT
	eToManual		: E_ModeSwitch := E_ModeSwitch.Standby;	// Auto → Manual 때 어디까지
	eToAuto			: E_ModeSwitch := E_ModeSwitch.Zero;		// Manual → Auto 때 어디까지
	tDelay			: TIME := T#400MS;						// 출력 0으로 둔 뒤 다음 단계까지
	bKeepOnRestart	: BOOL;		// FALSE(기본) = PMS가 다시 켜지면 모든 유닛을 Manual로 시작 (요청 모드도 Manual로 씀. 정전 뒤 장비 투입은 운전원이 확인하고 함). TRUE = 저장된 요청 모드를 그대로 씀
END_STRUCT
END_TYPE

// ---- 10_Core/40_Arbitration/E_ModeSwitch.TcDUT
{attribute 'qualified_only'}
{attribute 'strict'}
TYPE E_ModeSwitch :		// 모드 전환 때 어디까지 하고 바꾸나
(
	Direct		:= 0,	// 바로 바꿈
	Zero		:= 1,	// 출력 0 → 지연 → 바꿈
	Standby		:= 2	// 출력 0 → 지연 → Standby (운전 중일 때만) → Run이 아니게 되면 바꿈
) INT;
END_TYPE

// ---- 10_Core/40_Arbitration/E_ModeStep.TcDUT
{attribute 'qualified_only'}
{attribute 'strict'}
TYPE E_ModeStep :
(
	Idle		:= 0,	// 전환 없음
	Zero		:= 1,	// 출력 0, 지연 중
	WaitStop	:= 2	// Standby 보냄, Run이 아니게 되기를 기다림
) INT;
END_TYPE

// ---- 10_Core/40_Arbitration/E_CmdRefuse.TcDUT
{attribute 'qualified_only'}
{attribute 'strict'}
TYPE E_CmdRefuse :		// 무시한 지령의 이유
(
	None		:= 0,
	Reversed	:= 1	// Manual: 지금 출력 방향과 반대
) INT;
END_TYPE

// ---- 10_Core/50_Distribution/ST_UnitDiag.TcDUT
TYPE ST_UnitDiag :
STRUCT
	eRole		: E_UnitRole;
	fPReq		: REAL;				// kW, 그룹 안에서 나눈 직후 값 (배터리·S 확인 전)
	fPOut		: REAL;				// kW, 최종
	ePBy	: E_UnitLimitBy;	// P를 마지막으로 줄인 것
	nPModule	: UINT;	// P를 줄인 모듈 (유닛 제한·버스 제한 모듈). 0 = 코어
	fQReq		: REAL;
	fQOut		: REAL;
	eQBy		: E_UnitLimitBy;
	(* 따라가기용 중간값 (P) *)
	fPMax	: REAL;	// kW, 유닛 한도 = 설비 한도 (FB_EquipmentLimits. 운전 대상 아니면 0)
	fPWeight	: REAL;				// 그룹 몫을 나눌 때 쓴 무게 (분배 기준: 정격·SOC·균등)
	fPBat		: REAL;				// kW, 배터리 그룹 방향·한도 적용 후 (피상전력 전)
END_STRUCT
END_TYPE

// ---- 10_Core/50_Distribution/ST_DistDiag.TcDUT
TYPE ST_DistDiag :		// 분배 진단 (그룹 하나): Manual을 먼저 나누고, Auto는 Manual이 덜 나간 만큼 더해서 나눔
STRUCT
	stAutoP		: ST_DistPathDiag;		// kW
	stManualP	: ST_DistPathDiag;
	stAutoQ		: ST_DistPathDiag;		// kvar
	stManualQ	: ST_DistPathDiag;
END_STRUCT
END_TYPE

// ---- 10_Core/50_Distribution/ST_DistPathDiag.TcDUT
TYPE ST_DistPathDiag :		// 분배 진단: 경로(Auto 또는 Manual) 하나, P 또는 Q 하나
STRUCT
	fTarget		: REAL;		// 이 경로 목표 (Auto는 Manual이 덜 나간 만큼 더한 값)
	fFixed		: REAL;		// 유닛별 값 합 (유닛 한도 후, 축소 전)
	fShareReq	: REAL;		// 그룹 몫 유닛에 나눠야 할 양 (방향 규칙 후). 그룹 지령 없으면 0
	fShareGot	: REAL;		// 실제로 나눈 양 (유닛 한도 때문에 작을 수 있음)
	fFixedScale	: REAL;		// 유닛별 값 축소 비율 (1 = 안 줄임)
	fOut		: REAL;		// 이 경로 유닛 합 (배터리 버스·피상전력 전)
END_STRUCT
END_TYPE

// ---- 10_Core/50_Distribution/ST_BatDistDiag.TcDUT
TYPE ST_BatDistDiag :		// 배터리 그룹(DC 버스)별 분배 따라가기
STRUCT
	fNetIn		: REAL;		// kW, 그룹 분배 직후 이 버스 유닛 P 합
	nDirZero	: UINT;		// 순 방향과 반대라 0으로 만든 유닛 수
	fNetDir		: REAL;		// kW, 방향 맞춘 뒤 합
	fLimit		: REAL;		// kW, 그 방향 한도 (방전 +, 충전 -)
	fScale		: REAL;		// 한도 때문에 곱한 비율 (1 = 안 줄임)
END_STRUCT
END_TYPE

// ---- 10_Core/00_Type/E_SelectMode.TcDUT
{attribute 'qualified_only'}
{attribute 'strict'}
TYPE E_SelectMode :
(
	Grade		:= 0,	// 등급 우선 (등급 숫자가 작은 지령원)
	MinAbs		:= 1	// 절대값이 가장 작은 값
) INT;
END_TYPE

// ---- 10_Core/00_Type/ST_GroupSet.TcDUT
TYPE ST_GroupSet :
STRUCT
	eSelP		: E_SelectMode;		// 그룹 P 지령원 고르는 방식
	eSelQ		: E_SelectMode;		// 그룹 Q 지령원 고르는 방식
	bRamp		: BOOL;				// 램프 사용 (Auto·Manual 공통). FALSE = 램프율과 관계없이 바로 목표 (기본)
	fRampUp		: REAL;				// kW/s, |P|가 커지는 쪽. 0 = 램프 없음
	fRampDn		: REAL;				// kW/s, |P|가 작아지는 쪽. 0 = 램프 없음
	fRampResume	: REAL;				// kW/s, 제한 모듈이 재개 중일 때 오르는 쪽. 0 = fRampUp 사용
	tQFilter	: TIME;				// Q 응답 필터 시정수. T#0S = 필터 없음
	eDistBasis	: E_DistBasis := E_DistBasis.Soc;	// 그룹 몫 나누는 기준. 기본 SOC (방전은 SOC 높은 쪽, 충전은 낮은 쪽이 많이. Q는 정격 비율). 현장에서 다른 기준을 쓰려면 GVL_PERSIST.g_astGroupSet 초기값에서
	bQPriority	: BOOL;				// 피상전력 초과 시 TRUE = Q 우선, FALSE = P 우선
END_STRUCT
END_TYPE

// ---- 10_Core/00_Type/ST_ManualPolicy.TcDUT
TYPE ST_ManualPolicy :		// 제어 그룹마다 Manual 경로에 적용할 단계 (TRUE = 적용). Auto 경로는 항상 전부 적용
STRUCT
	(* 운전 정책 *)
	bRamp		: BOOL := TRUE;		// P 램프·Q 응답 필터 (그룹 설정 bRamp·tQFilter를 따름)
	bSrcLimit	: BOOL := TRUE;		// 지령원이 낸 P 제한
	bPccLimit	: BOOL := TRUE;		// 접속점 기준 제한 모듈 (모듈 등록의 bManual = TRUE인 것만)
	bComp		: BOOL := FALSE;	// 보정 (같은 그룹에 Auto 유닛이 있으면 Auto 쪽에만 더함: 두 번 더하지 않게)
	bDevLimit	: BOOL := TRUE;		// 설비 기준 제한 모듈 (P·Q)
	(* 장비 한도 — 끄면 이 그룹 Manual 유닛은 PMS가 이 한도로 막지 않음 (장비 자체 보호는 그대로) *)
	bRating		: BOOL := TRUE;		// 유닛 정격·Derate·피상전력
	bBatLimit	: BOOL := TRUE;		// BMS 충방전 한도 (유닛·배터리 버스)
	(* 보호는 보호 항목마다 ST_ProtCfg.bManual로 켜고 끔 *)
END_STRUCT
END_TYPE

// ---- 10_Core/40_Arbitration/E_UnitRole.TcDUT
{attribute 'qualified_only'}
{attribute 'strict'}
TYPE E_UnitRole :
(
	None			:= 0,
	Fixed			:= 1,	// 유닛별 값을 따름
	AutoShare		:= 2,	// Auto 그룹 몫을 받음
	ManualShare		:= 3	// Manual 그룹 몫을 받음
) INT;
END_TYPE

// ---- 10_Core/40_Arbitration/ST_Pick.TcDUT
TYPE ST_Pick :
STRUCT
	bActive		: BOOL;		// 고른 값이 있음
	fValue		: REAL;		// kW 또는 kvar
	nModule		: UINT;		// 고른 지령원 모듈 ID
	bNew		: BOOL;		// 고른 지령원이 이번 스캔에 새 지령을 냄
END_STRUCT
END_TYPE

// ---- 10_Core/40_Arbitration/ST_Range.TcDUT
TYPE ST_Range :
STRUCT
	fMax		: REAL;		// 상한
	fMin		: REAL;		// 하한
	nMaxModule	: UINT;		// 상한을 정한 모듈 (0 = 코어)
	nMaxReason	: UINT;
	nMinModule	: UINT;		// 하한을 정한 모듈
	nMinReason	: UINT;
END_STRUCT
END_TYPE

// ---- 10_Core/40_Arbitration/ST_Clamp.TcDUT
TYPE ST_Clamp :
STRUCT
	fIn			: REAL;
	fOut		: REAL;
	bClamped	: BOOL;		// 값이 잘림
	nModule		: UINT;		// 자른 모듈 (0 = 코어)
	nReason		: UINT;
END_STRUCT
END_TYPE

// ---- 10_Core/40_Arbitration/ST_ShapeDiag.TcDUT
TYPE ST_ShapeDiag :		// 성형 진단: 경로(Auto 또는 Manual) 하나, 그룹 하나. 두 경로가 같은 모양
STRUCT
	(* P *)
	bPGroupCmd	: BOOL;			// 이 경로 그룹 P 지령 있음. 없으면 이 경로 유닛 지령 합이 목표 (지령 없는 유닛은 0)
	bPUnitCmd	: BOOL;			// 이 경로 유닛 P 지령이 하나라도 있음
	nPSource	: UINT;			// 고른 그룹 지령원 모듈 ID (0 = 그룹 지령 없음)
	fPReq		: REAL;			// kW, 그룹 지령 또는 유닛 지령 합 (램프 전)
	fPRamped	: REAL;			// kW, 램프 후 (유닛 지령 합이면 유닛별 램프 후 합)
	stPcc		: ST_Clamp;		// 접속점 제한 (지령원 P 제한 + 접속점 기준 모듈)
	fPComp		: REAL;			// kW, 더한 보정 합
	stDev		: ST_Clamp;		// 설비 제한 (보정 후: 가용 정격 + 배터리 한도 + 설비 기준 모듈)
	fPOut		: REAL;			// kW, 이 경로 몫 (Auto는 그룹 전체 목표에서 Manual 몫을 뺀 값)
	(* Q *)
	bQGroupCmd	: BOOL;
	bQUnitCmd	: BOOL;
	stQ			: ST_Clamp;
	(* 따라가기용 중간값 *)
	fRampUp		: REAL;			// kW/s, 이번 스캔에 쓴 오르기 램프율 (0 = 램프 없음, 재개 램프 포함)
	fRampDn		: REAL;			// kW/s, 내리기 램프율
	stPccRng	: ST_Range;		// P 접속점 제한 범위
	stDevRng	: ST_Range;		// P 설비 제한 범위
	stQRng		: ST_Range;		// Q 제한 범위
	stTrace		: ST_PTrace;	// P 추적표 (요청 → … → 설비 제한). 유닛 한도·분배와 쓴 값은 FB_OutputDiag가 덧붙임
END_STRUCT
END_TYPE

// ---- 10_Core/00_Type/ST_UnitReq.TcDUT
TYPE ST_UnitReq :
STRUCT
	bPSetActive	: BOOL;
	fPSet		: REAL;		// kW, 유닛 출력
	bQSetActive	: BOOL;
	fQSet		: REAL;		// kvar
END_STRUCT
END_TYPE

// ---- 10_Core/00_Type/ST_BmsCfg.TcDUT
TYPE ST_BmsCfg :
STRUCT
	nBatGroup	: UINT := 1;		// 소속 배터리 그룹(DC 버스). 유닛은 UNIT_CFG.nBatGroup으로 같은 그룹을 가리킴
	fCapacity	: REAL;				// kWh. SOC 가중 평균의 무게 (0 = 설정 안 함 → 무게 1)
END_STRUCT
END_TYPE

// ---- 10_Core/20_Protection/ST_BmsProt.TcDUT
TYPE ST_BmsProt :
STRUCT
	eBatAction	: E_BatAction;		// 이 BMS에 걸린 가장 센 조치
	nModule		: UINT;				// 조치를 건 보호 모듈 ID
END_STRUCT
END_TYPE

// ---- 10_Core/20_Protection/ST_BmsAvail.TcDUT
TYPE ST_BmsAvail :
STRUCT
	bUsable		: BOOL;		// 쓸 수 있음 (아래 이유가 하나도 없음)
	bNotInstalled	: BOOL;		// 미설치: BMS 칸이 비어 있음. 배터리 그룹 집계·보호에서 뺌
	bNoComm		: BOOL;
	bFault		: BOOL;
	bSysStop	: BOOL;		// BMS가 스스로 정지
	bProt		: BOOL;		// 배터리 보호 조치 중
END_STRUCT
END_TYPE

// ---- 10_Core/20_Protection/ST_BatGroupState.TcDUT
TYPE ST_BatGroupState :
STRUCT
	bUsable		: BOOL;		// 쓸 수 있는 BMS가 하나 이상
	bReady		: BOOL;		// 투입 완료: 쓸 수 있는 BMS가 하나 이상이고 전부 투입됨
	nBms		: UINT;		// 소속 BMS 수 (설치된 것만)
	nBmsUsable	: UINT;		// 쓸 수 있는 BMS 수
	fPChgMax	: REAL;		// kW, 쓸 수 있는 BMS 충전 한도 합 (양수)
	fPDisMax	: REAL;		// kW, 방전 한도 합
	stSoc		: ST_Val;	// %, 용량 가중 평균
	stSocMin	: ST_Val;	// %
	stSocMax	: ST_Val;	// %
	fSocWeight	: REAL;		// 평균에 쓴 무게 합 (그룹끼리 다시 평균낼 때 씀)
	fCapacity	: REAL;		// kWh, SOC가 유효한 쓸 수 있는 BMS 용량 합 (BMS_CFG.fCapacity. 설정 안 하면 0)
END_STRUCT
END_TYPE

// ---- 10_Core/00_Type/E_PcsAction.TcDUT
{attribute 'qualified_only'}
{attribute 'strict'}
TYPE E_PcsAction :		// 보호 조치 (PCS)
(
	None		:= 0,	// 조치 없음 (알람만), 자동 해제
	Standby		:= 1,	// 대기 = 출력 0 (명령 없음: 가용 아님으로 출력에서 빠짐). 조건이 있는 동안만, 풀리면 다시 출력
	Stop		:= 2,	// 정지 명령. 조건이 풀려도 정지 유지 (다시 운전하려면 Run)
	EStop		:= 3	// 비상정지. 위와 같음
) INT;
END_TYPE

// ---- 10_Core/00_Type/E_BatAction.TcDUT
{attribute 'qualified_only'}
{attribute 'strict'}
TYPE E_BatAction :
(
	None		:= 0,	// 조치 없음
	Stop		:= 1,	// 정지 (접촉기 개방). 잠금 없음. 다시 투입하려면 새 기동·투입 요청 필요
	EStop		:= 2	// 비상정지. 재투입 조건은 Stop과 같음
) INT;
END_TYPE

// ---- 10_Core/00_Type/E_ModeAction.TcDUT
{attribute 'qualified_only'}
{attribute 'strict'}
TYPE E_ModeAction :		// 보호가 운전 모드를 바꾸는가 (보호 항목마다 ST_ProtCfg.eModeAction)
(
	None		:= 0,	// 모드를 바꾸지 않음 (기본)
	ToManual	:= 1	// 조치를 받는 Auto 유닛의 요청 모드를 Manual로 바꿈. 보호가 풀려도 Manual 유지, 운전원이 Auto를 다시 요청
) INT;
END_TYPE

// ---- 10_Core/00_Type/ST_ProtCfg.TcDUT
TYPE ST_ProtCfg :
STRUCT
	bAuto		: BOOL := TRUE;		// Auto 유닛에 조치를 걸음
	bManual		: BOOL := TRUE;		// Manual 유닛에 조치를 걸음
	// 둘 중 하나라도 TRUE면 감지·발생 표시·로그. 둘 다 FALSE면 이 보호를 안 씀
	// 아래는 표준 대응(g_fbProtRespStd를 대응 칸에 등록)이 쓰는 조치. 대응 칸이 비면 조치 없음 (알람만, 문구도 조치 없음). 다른 대응 모듈을 붙이면 그 모듈이 정함
	// [결함 8 수정 2026-11-03: 주석 고침. 원래 '아래는 표준 대응(대응 칸이 비었을 때)이 쓰는 조치. 대응 모듈을 붙이면 그 모듈이 정함']
	// BMS 조치는 같은 버스에 조치를 받는 유닛이 하나라도 있을 때 (버스에 유닛이 없으면 그대로 걸음)
	ePcsAction	: E_PcsAction;		// PCS 조치: Standby = 출력 0 (명령 없음), Stop·EStop = 명령
	eBatAction	: E_BatAction;		// 배터리 조치. PCS가 Stop·EStop일 때만 고를 수 있음 (시퀀서가 버스 PCS 정지 확인 뒤 보냄)
	eModeAction	: E_ModeAction;		// 운전 모드 조치. ToManual = 조치를 받는 Auto 유닛의 요청 모드를 Manual로 바꿈 (보호가 풀려도 Manual 유지)
	fPPct		: REAL := 100.0;	// P 상한 (유닛 정격 대비 %). 100 = 줄이지 않음
	fQPct		: REAL := 100.0;	// Q 상한 (유닛 정격 대비 %). 100 = 줄이지 않음
END_STRUCT
END_TYPE

// ---- 10_Core/20_Protection/ST_UnitProt.TcDUT
TYPE ST_UnitProt :
STRUCT
	ePcsAction		: E_PcsAction;		// 이 유닛에 걸린 가장 센 조치
	nModule			: UINT;				// 조치를 건 보호 모듈 ID
	fPPct			: REAL := 100.0;	// 걸린 P 상한 중 가장 낮은 값 (유닛 정격 대비 %, 100 = 없음)
	nPModule		: UINT;			// P 상한을 건 모듈 ID
	fQPct			: REAL := 100.0;	// 걸린 Q 상한 중 가장 낮은 값 (유닛 정격 대비 %, 100 = 없음)
	nQModule		: UINT;			// Q 상한을 건 모듈 ID
	bModeManualReq	: BOOL;				// 보호가 걸려 있는 동안 TRUE: 이 유닛의 요청 모드를 Manual로 (실제 모드와 관계없음. FB_ModeSwitch가 요청값을 씀)
	nModeModule		: UINT;				// 모드 조치를 건 보호 모듈 ID
END_STRUCT
END_TYPE

// ---- 10_Core/20_Protection/ST_UnitAvail.TcDUT
TYPE ST_UnitAvail :
STRUCT
	bAvail		: BOOL;		// 출력 가능 (아래 이유가 하나도 없음). Derate는 가용에 영향 없음
	bNotInstalled	: BOOL;		// 미설치: 유닛의 PCS 칸이 비어 있음 (모니터링 전용 등). 통신·고장 판단·보호에서 뺌
	bNoPcsComm	: BOOL;
	bPcsFault	: BOOL;
	bPcsLocal	: BOOL;		// PCS가 PMS 제어를 안 받는 상태
	bNoBat		: BOOL;		// 연결 배터리 그룹에 쓸 수 있는 BMS가 없음 (그룹 번호 설정 오류 포함) → FB_BatGroup 결과에서 이유 확인
	bProt		: BOOL;		// 유닛 보호 조치 중 (대기·정지·비상정지)
END_STRUCT
END_TYPE

// ---- 10_Core/00_Type/ST_PointTerm.TcDUT
TYPE ST_PointTerm :
STRUCT
	nMeter		: UINT;				// 계측기 (GVL_SITE.g_aipMeter 칸). 0 = 빈 칸
	fSign		: REAL := 1.0;		// +1 더함, -1 뺌
END_STRUCT
END_TYPE

// ---- 10_Core/00_Type/ST_PointCfg.TcDUT
TYPE ST_PointCfg :		// 계측점 = 계측기 값을 부호와 함께 더한 것. 전압·주파수는 첫 계측기 값
STRUCT
	astTerm		: ARRAY[1..GVL_PARAM.POINT_TERM_MAX] OF ST_PointTerm;
END_STRUCT
END_TYPE

// ---- 10_Core/10_Snapshot/ST_VirtualSet.TcDUT
TYPE ST_VirtualSet :
STRUCT
	bVEna		: BOOL;		// 가상 전압 사용
	fV			: REAL;		// V, 상전압 (평균·A·B·C 모두 이 값)
	bPEna		: BOOL;		// 가상 유효전력 사용
	fP			: REAL;		// kW
END_STRUCT
END_TYPE

// ---- 10_Core/00_Type/E_GroupState.TcDUT
{attribute 'qualified_only'}
{attribute 'strict'}
TYPE E_GroupState :
(
	Init			:= 0,	// 부팅 직후: 첫 스냅샷 대기, 쓰기 금지
	Stopped			:= 1,
	BatConnecting	:= 2,	// 배터리 투입 확인
	PcsStandby		:= 3,	// PCS 대기 (활성 + 출력 0)
	StartWait		:= 4,	// 기동 조건(I_StartPermit) 대기. 등록된 조건이 없으면 바로 통과
	Running			:= 5,
	Stopping		:= 6	// 정지 램프 → 정지 명령 확인
) INT;
END_TYPE

// ---- 10_Core/00_Type/E_LimitBasis.TcDUT
{attribute 'qualified_only'}
{attribute 'strict'}
TYPE E_LimitBasis :
(
	Pcc			:= 0,	// 접속점 기준 (보정 전)
	Device		:= 1	// 설비 기준 (보정 후, PCS 출력 합)
) INT;
END_TYPE

// ---- 10_Core/00_Type/E_OpMode.TcDUT
{attribute 'qualified_only'}
{attribute 'strict'}
TYPE E_OpMode :
(
	Auto		:= 0,	// 자동: 원격·자동 지령원이 동작
	Manual		:= 1	// 수동: 수동 지령원만 동작
) INT;
END_TYPE

// ---- 10_Core/00_Type/E_ProtScope.TcDUT
{attribute 'qualified_only'}
{attribute 'strict'}
TYPE E_ProtScope :
(
	Unit		:= 0,	// 유닛 하나
	Bms			:= 1,	// BMS 하나 (PCS 조치는 그 BMS가 속한 배터리 그룹의 유닛에)
	BatGroup	:= 2,	// 배터리 그룹(DC 버스) 하나: 그 그룹의 BMS와 유닛 전부
	Group		:= 3,	// 제어 그룹 하나
	Site		:= 4	// 사이트 전체
) INT;
END_TYPE

// ---- 10_Core/00_Type/E_RunState.TcDUT
{attribute 'qualified_only'}
{attribute 'strict'}
TYPE E_RunState :
(
	Unknown		:= 0,	// 통신 전, 해석 불가
	Stop		:= 1,
	Standby		:= 2,	// 대기: 활성인데 출력 0 (Total Interface 대기)
	Run			:= 3,	// 활성: 출력 지령을 받음 (크기 무관)
	Fault		:= 4
) INT;
END_TYPE

// ---- 10_Core/00_Type/E_SourceMode.TcDUT
{attribute 'qualified_only'}
{attribute 'strict'}
TYPE E_SourceMode :
(
	Auto		:= 0,	// 자동 모드에서만 동작
	Manual		:= 1,	// 수동 모드에서만 동작
	Both		:= 2,	// 운전 모드와 관계없이 동작
	None		:= 3	// 받지 않음
) INT;
END_TYPE

// ---- 10_Core/00_Type/ST_BatState.TcDUT
TYPE ST_BatState :
STRUCT
	bComm			: BOOL;
	bContactorClosed: BOOL;
	bWarn			: BOOL;
	bFault			: BOOL;
	bSysStop		: BOOL;		// 배터리가 스스로 정지 (운전 불가)
	stSoc			: ST_Val;	// %
	stSoh			: ST_Val;	// %
	fPChgMax		: REAL;		// kW, 충전 한도 (양수). bComm = FALSE면 0으로 본다
	fPDisMax		: REAL;		// kW, 방전 한도 (양수)
	bWriteFail		: BOOL;		// 장비 쓰기(명령)가 잇달아 실패함 (드라이버가 FB_DeviceBase.M_MarkWriteResult로 판단해 채움)
END_STRUCT
END_TYPE

// ---- 10_Core/00_Type/ST_GroupCfg.TcDUT
TYPE ST_GroupCfg :
STRUCT
	nPccPoint	: UINT := 1;		// 접속점 계측점 (GVL_SITE.POINT_CFG 칸). 0 = 없음
END_STRUCT
END_TYPE

// ---- 10_Core/00_Type/ST_GroupView.TcDUT
TYPE ST_GroupView :
STRUCT
	nGroup			: UINT;				// 제어 그룹 번호
	eState			: E_GroupState;
	stPcc			: ST_PccMeas;		// 접속점 계측
	fPRatedSum		: REAL;				// kW, 그룹 유닛 정격 합 (가용과 관계없이 전부)
	fQRatedSum		: REAL;				// kvar
	nUnitAvail		: UINT;				// 가용 유닛 수
	fPRatedAvail	: REAL;	// kW, 가용 유닛 P 한도 합 (정격 × Derate ∩ 유닛 제한 모듈. FB_EquipmentLimits 그룹 정격 줄)
	fQRatedAvail	: REAL;	// kvar, 가용 유닛 Q 한도 합
	fSRatedAvail	: REAL;	// kVA, 가용 유닛 피상전력 한도 합
	fPChgMax	: REAL;	// kW, 배터리 기준 그룹 충전 한도 (양수. 버스 한도·버스 제한 모듈 반영, FB_EquipmentLimits 배터리 줄)
	fPDisMax	: REAL;	// kW, 배터리 기준 그룹 방전 한도 (양수)
	stSocMin		: ST_Val;			// %
	stSocMax		: ST_Val;			// %
	stSocAvg		: ST_Val;			// %
	fCapacity		: REAL;				// kWh, 가용 유닛이 쓰는 배터리 그룹 용량 합 (BMS_CFG.fCapacity. 0 = 설정 안 함)
	fPOut			: REAL;				// kW, 유닛 출력 합 (실측)
	fQOut			: REAL;				// kvar
END_STRUCT
END_TYPE

// ---- 10_Core/00_Type/ST_Limit.TcDUT
TYPE ST_Limit :
STRUCT
	bActive		: BOOL;
	fMax		: REAL;		// 상한 (방전·공급 쪽)
	fMin		: REAL;		// 하한 (충전·흡수 쪽)
	nModule		: UINT;		// 낸 모듈 ID. 0 = 코어
	nReason		: UINT;		// 모듈 안의 이유 코드. 0 = 없음
END_STRUCT
END_TYPE

// ---- 10_Core/00_Type/ST_LimitOut.TcDUT
TYPE ST_LimitOut :
STRUCT
	stP			: ST_Limit;	// kW
	stQ			: ST_Limit;	// kvar
	bResume		: BOOL;		// 출력 재개 중: 코어 램프가 재개 램프율을 쓴다
END_STRUCT
END_TYPE

// ---- 10_Core/00_Type/ST_MeterState.TcDUT
TYPE ST_MeterState :
STRUCT
	bComm		: BOOL;
	stP			: ST_Val;					// kW
	stQ			: ST_Val;					// kvar
	stV			: ST_Val;					// V, 상전압 평균
	astV		: ARRAY[1..3] OF ST_Val;	// V, A·B·C 상전압
	stF			: ST_Val;					// Hz
END_STRUCT
END_TYPE

// ---- 10_Core/00_Type/ST_ModuleReg.TcDUT
TYPE ST_ModuleReg :
STRUCT
	bEnable		: BOOL := TRUE;
	nGroup		: UINT;					// 대상 제어 그룹. 0 = 모든 그룹 (제한·보정·기동 조건은 그룹이 1개일 때만. 2개 이상이면 그룹마다 인스턴스)
	bManual		: BOOL := TRUE;			// 출력 제한 모듈만: 접속점 기준 모듈을 Manual 경로에도 적용 (Auto는 항상 적용). 기본 TRUE: 역송 방지·계약 전력처럼 넘으면 안 되는 상한은 Manual도 지킴. 현장 시험 때만 FALSE로 풀고 끝나면 TRUE (영속값이라 저절로 안 돌아옴)
	// [5-16 결정 2026-11-04: 기본값 TRUE로. 원래 bManual : BOOL; (기본 FALSE). 이미 운영 중인 현장은 저장된 값(FALSE)이 그대로 남으므로 업데이트 때 TRUE로 한 번 씀]
END_STRUCT
END_TYPE

// ---- 10_Core/00_Type/ST_PQ.TcDUT
TYPE ST_PQ :		// P·Q 한 쌍 (유닛 지령·쓴 값·보정량 공통)
STRUCT
	fP			: REAL;		// kW, 방전·공급 +
	fQ			: REAL;		// kvar, 공급 +
END_STRUCT
END_TYPE

// ---- 10_Core/00_Type/ST_PccMeas.TcDUT
TYPE ST_PccMeas :
STRUCT
	stMeas		: ST_MeterState;	// 제어용 값 (가상신호 적용 후)
	bNoPoint	: BOOL;				// 접속점 계측점이 없음 (GROUP_CFG.nPccPoint 0 = 없음). [결함 7 수정 2026-11-03: 추가]
END_STRUCT
END_TYPE

// ---- 10_Core/00_Type/ST_RuleCfg.TcDUT
TYPE ST_RuleCfg :		// 현장 보호 규칙(모듈) 하나의 설정
STRUCT
	stProt		: ST_ProtCfg;			// 사용 모드 (bAuto·bManual)·표준 대응 조치
	eScope		: E_ProtScope;			// Unit / Bms / BatGroup / Group / Site
	nTarget		: UINT;					// 대상 번호 (유닛·배터리 그룹·제어 그룹). Site면 무시
	fThreshold	: REAL;					// 임계값 (단위는 규칙마다)
END_STRUCT
END_TYPE

// ---- 10_Core/00_Type/ST_SourceOutput.TcDUT
TYPE ST_SourceOutput :
STRUCT
	bValid			: BOOL;			// 사용 중 + 유효 + 만료 안 됨. FALSE면 아래 전부 무시
	(* P 지령 *)
	bPSetActive		: BOOL;
	fPSet			: REAL;			// kW, 접속점 기준
	(* P 제한 *)
	bPLimActive		: BOOL;
	fPMax			: REAL;			// kW
	fPMin			: REAL;			// kW
	(* Q 지령 *)
	bQSetActive		: BOOL;
	fQSet			: REAL;			// kvar, 접속점 기준
	(* Q 제한 *)
	bQLimActive		: BOOL;
	fQMax			: REAL;			// kvar, 공급 상한 (접속점 기준)
	fQMin			: REAL;			// kvar, 흡수 하한
	bNewSet			: BOOL;			// 새 지령값이 들어옴 (1스캔). Manual 유닛은 이 스캔에 바로 씀
	(* 상태 요청 *)
	stPcsReq		: ST_PcsReq;		// PCS 상태 요청 (Run·Standby·Stop·EStop·Reset)
	stBatReq		: ST_BatReq;		// 배터리 요청 (Close·Open)
	(* 유닛별 값 (선택) *)
	astUnit			: ARRAY[1..GVL_PARAM.UNIT_COUNT] OF ST_UnitReq;	// 값이 있는 유닛은 그룹 몫 대신 이 값
END_STRUCT
END_TYPE

// ---- 10_Core/00_Type/ST_SourceReg.TcDUT
TYPE ST_SourceReg :
STRUCT
	bEnable		: BOOL;
	nGrade		: UINT := 9;			// 등급. 1이 가장 높음
	stStateMode	: ST_StateModeSet;					// 상태 요청을 명령마다 어느 운전 모드에서 받나 (기본 모두 Manual). 리셋은 모드와 관계없이 받음
	ePowerMode	: E_SourceMode := E_SourceMode.Auto;	// P·Q 지령과 P 제한을 받는 운전 모드
	nGroup		: UINT;					// 대상 제어 그룹. 0 = 모든 그룹
	tExpire		: TIME := T#10S;		// 이 시간 동안 새 값이 없으면 끊김
	bLostAlarm	: BOOL := TRUE;			// 끊기면 '지령원 끊김' 알람 (FB_EventLog). FALSE = 알람 안 냄 (끊김 처리는 그대로). [9번 수정 2026-11-09: 추가 — EMS는 브로커 끊김 알람으로 대신]
END_STRUCT
END_TYPE

// ---- 10_Core/00_Type/E_PcsCmd.TcDUT
{attribute 'qualified_only'}
{attribute 'strict'}
TYPE E_PcsCmd :		// PCS(유닛) 상태 명령
(
	None		:= 0,
	Run			:= 1,	// 활성 (정지면 기동)
	Standby		:= 2,	// 대기 = 활성 + 출력 0 (정지면 기동 후 대기)
	Stop		:= 3,
	Reset		:= 4,	// 고장 리셋: 그 장비에 고장 리셋 명령 (PMS 상태는 바꾸지 않음)
	EStop		:= 5	// 비상정지
) INT;
END_TYPE

// ---- 10_Core/00_Type/E_BatCmd.TcDUT
{attribute 'qualified_only'}
{attribute 'strict'}
TYPE E_BatCmd :		// 배터리(BMS) 명령
(
	None		:= 0,
	Close		:= 1,	// DC 접촉기 투입
	Open		:= 2,	// DC 접촉기 개방
	EStop		:= 3,	// 비상정지 (보호)
	Reset		:= 4	// 고장 리셋
) INT;
END_TYPE

// ---- 10_Core/00_Type/ST_PcsCmd.TcDUT
TYPE ST_PcsCmd :		// PCS(유닛)에 보낼 명령
STRUCT
	eCmd		: E_PcsCmd;
	nSeq		: UDINT;		// 명령 번호. 바뀌면 새 명령 → 디스패처가 1회 전송
END_STRUCT
END_TYPE

// ---- 10_Core/00_Type/ST_BatCmd.TcDUT
TYPE ST_BatCmd :		// BMS에 보낼 명령
STRUCT
	eCmd		: E_BatCmd;
	nSeq		: UDINT;		// 명령 번호. 바뀌면 새 명령 → 디스패처가 1회 전송
END_STRUCT
END_TYPE

// ---- 10_Core/00_Type/ST_PcsReq.TcDUT
TYPE ST_PcsReq :		// 지령원의 PCS 상태 요청
STRUCT
	eCmd		: E_PcsCmd;		// None = 요청 없음. 새 요청일 때 1스캔만
	nUnit		: UINT;			// 대상 유닛. 0 = 지령원 대상 그룹 전체
END_STRUCT
END_TYPE

// ---- 10_Core/00_Type/ST_BatReq.TcDUT
TYPE ST_BatReq :		// 지령원의 배터리 요청
STRUCT
	eCmd		: E_BatCmd;		// Close / Open만 씀. None = 요청 없음. 새 요청일 때 1스캔만
	nBatGroup	: UINT;			// 대상 배터리 그룹. 0 = 전체
END_STRUCT
END_TYPE

// ---- 10_Core/00_Type/ST_PcsSeqSet.TcDUT
TYPE ST_PcsSeqSet :		// PCS(유닛) 시퀀스 설정
STRUCT
	tCmdConfirm		: TIME := T#30S;		// 기동 쪽 명령(Run) 접수 확인 시간. 지나면 실패 알람 (재시도 없음)
	tStopRetry		: TIME := T#5S;			// 정지 쪽 명령(Stop·EStop) 확인 시간·재시도 간격
	nStopRetry		: UINT := 3;			// 보호 명령(정지 쪽) 재시도 횟수. 넘으면 실패 알람만 (잠그지 않음)
	// 지령원 명령(운전원·EMS)은 운전 모드와 관계없이 재시도하지 않음: 한 번만 보내고, 확인 시간이 지나면 명령 실패 기록
	bStopRamp		: BOOL;					// 정지 전에 출력을 0까지 내림 (기본: 바로 Stop)
	fStopDonePct	: REAL := 1.0;			// 정지 램프 완료: |P| ≤ 유닛 정격의 이 %
	tStopRampMax	: TIME := T#30S;		// 정지 램프 최대 대기. 지나면 그대로 Stop
END_STRUCT
END_TYPE

// ---- 10_Core/00_Type/ST_BatSeqSet.TcDUT
TYPE ST_BatSeqSet :		// 배터리 시퀀스 설정
STRUCT
	eClose			: E_BatClose;			// 투입 시점 (OnStart / OnRequest). 새 기동·요청이 있어야 투입 (보호·고장으로 열린 뒤 저절로 다시 넣지 않음)
	bOpenOnStop		: BOOL;					// 버스의 유닛이 모두 정지하면 개방 (기본: 투입 유지)
	tConfirm		: TIME := T#60S;		// 투입 확인 시간. 지나면 실패 알람 (재시도 없음)
	tOpenRetry		: TIME := T#5S;			// 개방·비상정지 확인 시간·재시도 간격
	nOpenRetry		: UINT := 3;			// 보호 조치(개방·비상정지) 재시도 횟수. 넘으면 실패 알람만 (잠그지 않음)
	// 보호 조치가 아닌 명령(지령원 요청·자동 투입·정지 시 개방)은 한 번만 보냄
END_STRUCT
END_TYPE

// ---- 10_Core/00_Type/ST_ManualCmdSet.TcDUT
TYPE ST_ManualCmdSet :		// Manual 지령 거르기 설정 (FB_GateManual). 켜고 끔
STRUCT
	(* 1) Manual 방향 반대 지령 무시 (충전 중 방전, 방전 중 충전). 앞 값 유지 *)
	bReverse		: BOOL := TRUE;
	fDirBand		: REAL := 1.0;			// %, 실제 |P|가 정격의 이 % 이하면 멈춘 것으로 봄
	(* 2) Manual 지령은 Run을 확인한 뒤 들어온 것만 씀. Run이 아니거나 Manual로 막 바뀌면 새 지령이 올 때까지 0 *)
	bClearOnStop	: BOOL := TRUE;
	(* 배터리 한계는 버스 제한 모듈 (FB_SocLimit, GVL_SITE) *)
END_STRUCT
END_TYPE

// ---- 10_Core/00_Type/ST_StateModeSet.TcDUT
TYPE ST_StateModeSet :		// 지령원의 상태 요청을 명령마다 어느 운전 모드에서 받나 (Auto / Manual / Both / None). 리셋은 항상 받음
STRUCT
	stPcs		: ST_PcsCmdMode;	// PCS(유닛): Run·Standby·Stop·EStop
	stBat		: ST_BatCmdMode;	// 배터리 그룹: 투입·개방
END_STRUCT
END_TYPE

// ---- 10_Core/00_Type/ST_PcsCmdMode.TcDUT
TYPE ST_PcsCmdMode :		// PCS(유닛) 상태 요청을 명령마다 어느 운전 모드에서 받나 (기본 Manual: Auto에서는 지령원 상태 요청을 받지 않음. 보호·코어 요청은 모드와 관계없음)
STRUCT
	eRun		: E_SourceMode := E_SourceMode.Manual;	// Run
	eStandby	: E_SourceMode := E_SourceMode.Manual;	// Standby
	eStop		: E_SourceMode := E_SourceMode.Manual;	// Stop
	eEStop		: E_SourceMode := E_SourceMode.Manual;	// 비상정지
END_STRUCT
END_TYPE

// ---- 10_Core/00_Type/ST_BatCmdMode.TcDUT
TYPE ST_BatCmdMode :		// 배터리(배터리 그룹) 요청을 명령마다 어느 운전 모드에서 받나 (기본 Manual)
STRUCT
	eClose		: E_SourceMode := E_SourceMode.Manual;	// 배터리 투입
	eOpen		: E_SourceMode := E_SourceMode.Manual;	// 배터리 개방
END_STRUCT
END_TYPE

// ---- 10_Core/00_Type/ST_UnitCfg.TcDUT
TYPE ST_UnitCfg :
STRUCT
	nPcs		: UINT := 1;		// 소속 PCS 번호 (GVL_SITE.g_aipPcs 칸)
	nSub		: UINT := 1;		// PCS 안의 유닛 번호 (1..GVL_PARAM.MAX_SUB)
	nBatGroup	: UINT := 1;		// 연결된 배터리 그룹(DC 버스). BMS는 BMS_CFG.nBatGroup으로 같은 그룹에 속함. 0 = 연결 없음
	nGroup		: UINT := 1;		// 소속 제어 그룹
	fPRated		: REAL;				// kW
	fQRated		: REAL;				// kvar
	fSRated		: REAL;				// kVA
END_STRUCT
END_TYPE

// ---- 10_Core/00_Type/ST_UnitState.TcDUT
TYPE ST_UnitState :
STRUCT
	bComm		: BOOL;			// 통신 정상
	eRunState	: E_RunState;
	bCtrlReady	: BOOL := TRUE;	// PMS 제어를 받을 수 있는 상태 (리모트). 리모트 신호가 없는 장비는 드라이버가 건드리지 않음 → 리모트로 봄
	bFault		: BOOL;
	bWriteFail	: BOOL;			// 장비 쓰기(명령·지령)가 잇달아 실패함 (드라이버가 FB_DeviceBase.M_MarkWriteResult로 판단해 채움)
	stP			: ST_Val;		// kW
	stQ			: ST_Val;		// kvar
	eGridMode	: E_GridMode := E_GridMode.Gfl;	// 계통 제어 방식 (드라이버가 채움, 화면·로그용). 모르는 장비는 드라이버가 건드리지 않음 → GFL로 봄
END_STRUCT
END_TYPE

// ---- 10_Core/00_Type/ST_Val.TcDUT
TYPE ST_Val :
STRUCT
	fValue		: REAL;
	bValid		: BOOL;		// FALSE면 fValue를 쓰지 않는다
END_STRUCT
END_TYPE

// ---- 10_Core/00_Type/ST_OutputCfg.TcDUT
TYPE ST_OutputCfg :		// 출력 규칙 설정 (칸 번호 = GVL_SITE.g_aipOutput 칸)
STRUCT
	bEnable		: BOOL;
	nAux		: UINT;			// 낼 보조 장비 칸 (GVL_SITE.g_aipAux). 0 = 판단만 하고 안 냄
	nPoint		: UINT;			// 그 장비의 디지털 출력 점 번호
	fThreshold	: REAL;			// 규칙에 넘기는 값 (예: 팬 켜는 온도)
	tOnDelay	: TIME;			// 조건이 이 시간 유지되면 켬
	tOffDelay	: TIME;			// 조건이 없어지고 이 시간 뒤에 끔
	bLatch		: BOOL;			// 켜지면 리셋할 때까지 유지 (리셋은 조건이 없을 때만 풀림)
END_STRUCT
END_TYPE

// ---- 10_Core/00_Type/ST_ProtReq.TcDUT
TYPE ST_ProtReq :		// 보호 대응이 내는 요청 (보호 칸 하나·대상 하나). 코어가 대응을 부르기 전에 비우고, 부른 뒤 장비마다 합침 (센 쪽·낮은 쪽)
// 칸은 추가만 함 (새 칸의 기본값은 '요청 없음'이라 있던 대응 모듈은 그대로 동작)
STRUCT
	aePcs		: ARRAY[1..GVL_PARAM.UNIT_COUNT] OF E_PcsAction;		// 유닛 PCS 조치: Standby = 출력 0 (명령 없음), Stop·EStop = 명령
	abToManual	: ARRAY[1..GVL_PARAM.UNIT_COUNT] OF BOOL;			// 유닛 요청 모드를 Manual로 (걸려 있는 동안. 풀려도 Manual 유지)
	afPPct		: ARRAY[1..GVL_PARAM.UNIT_COUNT] OF REAL;	// 유닛 P 상한 (정격 대비 %, 100 = 없음. 코어가 비울 때 100으로 채움)
	afQPct		: ARRAY[1..GVL_PARAM.UNIT_COUNT] OF REAL;	// 유닛 Q 상한 (정격 대비 %, 100 = 없음. 코어가 비울 때 100으로 채움)
	aeBat		: ARRAY[1..GVL_PARAM.BMS_COUNT] OF E_BatAction;		// BMS 조치 (시퀀서가 버스 PCS 정지 확인 뒤 보냄)
END_STRUCT
END_TYPE

// ---- 10_Core/00_Type/ST_ProtView.TcDUT
TYPE ST_ProtView :		// 보호 모듈에 넘기는 정보 (대상 하나). 칸은 추가만 함 (이름 바꾸기·삭제 금지: 복사한 모듈이 깨짐)
STRUCT
	eScope		: E_ProtScope;		// 범위 (g_astRuleCfg.eScope)
	nTarget		: UINT;				// 지금 판단하는 대상 번호 (유닛·BMS·배터리 그룹·제어 그룹). Site면 1
	fThreshold	: REAL;				// 임계값 (g_astRuleCfg.fThreshold, 단위는 모듈마다)
	bInstalled	: BOOL;				// 대상 장비가 설치됨 (유닛 = PCS 칸, BMS = BMS 칸이 있음). 다른 범위는 TRUE
	(* 범위가 Unit일 때 *)
	stUnit		: ST_UnitState;		// 유닛 상태
	eOpMode		: E_OpMode;			// 유닛의 실제 운전 모드
	(* 범위가 Bms일 때 *)
	stBms		: ST_BatState;		// BMS 상태
	(* 범위가 Group일 때 *)
	stPcc		: ST_PccMeas;		// 접속점 계측
	(* 소속 (Unit: 그 유닛의 것, Bms: 그 BMS의 배터리 그룹, BatGroup·Group: 대상 번호) *)
	nGroup		: UINT;				// 제어 그룹
	nBatGroup	: UINT;				// 배터리 그룹 (0 = 배터리 없음)
END_STRUCT
END_TYPE

// ---- 20_Module/Mqtt/ST_MqttCommand_Rx.TcDUT
{attribute 'pack_mode' := '1'}
TYPE ST_MqttCommand_Rx :
STRUCT	// 인터페이스 100.Command 버전 2 (2026-11-25): 16 B, SequenceNumber 없음
	DeviceIndex	:	UDINT;	// 장치 번호 1부터 (F_MqttDistribute가 레코드 맨 앞에서 읽음: nIndexOffset = 0)
	CommandType	:	UDINT;
	Value		:	REAL;	// kW 등, CommandType에 따라 의미가 다름
	Delay		:	UDINT;	// ms. 이만큼 기다렸다가 실행 (0이면 바로). FB_EmsCmdGate
END_STRUCT
END_TYPE

// ---- 20_Module/Mqtt/ST_MqttCommandHeader.TcDUT
{attribute 'pack_mode' := '1'}
TYPE ST_MqttCommandHeader :
STRUCT
	HeaderVersion	:	UDINT;
	CommandVersion	:	UDINT;
	DeviceCount		:	UDINT;		// 이 메시지에 실린 장치 레코드 개수
	Location		:	UDINT;		// 0: PMS, 1: LOCAL, 2: CLOUD
	SiteID			:	UDINT;
	UserName		:	STRING(19);		//EMS에서 준 것 그대로 전송
	TimeStamp		:	STRING(23);
END_STRUCT
END_TYPE

// ---- 20_Module/Mqtt/ST_MqttHeader.TcDUT
{attribute 'pack_mode' := '1'}
TYPE ST_MqttHeader :
STRUCT
	HeaderVersion	:	UDINT;
	DeviceVersion	:	UDINT;
	SiteId			:	UDINT;
	DeviceCount		:	UDINT;		// 이 메시지에 실린 장치 레코드 개수
	TimeStamp		:	STRING(23);	// "2024-09-04 11:11:11.123" 형식 (23자 + null = 24byte)
END_STRUCT
END_TYPE

// ---- 20_Module/Mqtt/ST_MqttPubEntry.TcDUT
TYPE ST_MqttPubEntry :
STRUCT
	sTopic			:	STRING(30);	// device_name (예: 'pms', 'pcs', 'bat')
	pDeviceSrc		:	PVOID;			// 원본 장치 배열 시작 주소(매핑 완료된 wire-format 배열)
	nDeviceElemSize:	UDINT;			// 장치 레코드 1개 크기
	nDeviceCount	:	UDINT;			// 장치 개수 (헤더의 DeviceCount로도 사용)
	pStaging		:	PVOID;			// [헤더+장치배열] 조립용 스테이징 버퍼 시작 주소
	nStagingSize	:	UDINT;			// 스테이징 버퍼 전체 크기 (SIZEOF(Header) + 장치배열 크기)
	
	sCategory       : STRING(10);	//config전용  토픽 2번째 세그먼트. 'command' 또는 'config'
END_STRUCT
END_TYPE

// ---- 20_Module/Mqtt/ST_MqttSubEntry.TcDUT
TYPE ST_MqttSubEntry :
STRUCT
	sCategory		:	STRING(10);	// 토픽 2번째 세그먼트. 'command' 또는 'config'
	sTopic			:	STRING(20);	// device_name (예: 'pcs', 'bat', 'protection')
	bIndexed		:	BOOL;			// TRUE: 레코드 선두 DeviceIndex/DeviceId(UDINT)로 배열에 분배
									// FALSE: 헤더 뒤 레코드 1개를 목적지에 그대로 복사(고정 1건, protection 등)
	pDestArray		:	PVOID;			// 목적지 배열(또는 단일 구조체) 시작 주소
	nElementSize	:	UDINT;			// 레코드 1개 크기 (= 목적지 구조체 SIZEOF)
	nDeviceCapacity  : UDINT;//nMaxIndex		:	INT;			// bIndexed=TRUE일 때만 사용. 목적지 배열의 최대 인덱스(0-based)
	nSeqNum			:	UINT;			// 토픽별 수신 카운터. 100 초과 시 0으로 초기화

	pRxBuffer		:	PVOID;		// 이 토픽 전용 수신 버퍼 주소
	nRxBufferSize	:	UDINT;		// 그 버퍼의 실제 크기
	
	nMaxRecords      : UDINT;   // (nRxBufferSize - SIZEOF(Header)) / nElementSize, 빌드 시 1회 계산
	
	nDeviceIdBase	: UDINT;		// DEVICE_ID_BASE(1)에 더하는 토픽별 추가 시작 번호. 지금은 모두 0 [1부터 2026-11-10]
	nIndexOffset	: UDINT;		// 레코드 시작에서 DeviceIndex/DeviceId까지 바이트. 버전 2 command·config 모두 0 [2026-11-25]
END_STRUCT
END_TYPE
//dgsems/{solution}/{site_id}/{category}/{device_name}

// ---- 20_Module/Mqtt/Publish/ST_AirConditionerPublish_V1.TcDUT
(* 공조기(에어컨) 발행 레코드 1대 (명세: 21._Airconditioner.xlsx 시트 V1). 필드 이름·순서·형식은 명세 그대로 *)
{attribute 'pack_mode' := '1'}
TYPE ST_AirConditionerPublish_V1 :
STRUCT
	DeviceIndex			:	UDINT;		// 장치 인덱스
	Status				:	UDINT;		// 상태 (bit) b0 통신 이상, b1 정지, b2 운전, b3 알람
	ModeState			:	UDINT;		// 에어컨 모드 (enum) 0 Cooling, 2 Normal, 3 Auto, 4 Heating, 5 Dry, 6 Fan
	WindMode			:	UDINT;		// 바람 모드 (enum) 0 Normal, 1 Low, 2 Middle, 3 High, 4 Auto
	RoomTemperature		:	REAL;		// 실내 온도 ℃ (-1000 ~ 1000)
	ControlTemperature	:	REAL;		// 설정 온도 ℃ (-1000 ~ 1000)
	Fault1				:	UDINT;		// 고장 (bit) b0 실내 공기 온도 센서, b1 배관 입구 온도 센서, b2 유선 리모컨 통신, b3 Drain pump, b4 배관 출구 온도 센서, b5 EEPROM, b6 팬 Lock
END_STRUCT
END_TYPE

// ---- 20_Module/Mqtt/Publish/ST_BatPublish_V1.TcDUT
{attribute 'pack_mode' := '1'}
TYPE ST_BatPublish_V1 :
STRUCT
	DeviceIndex : UDINT; // 배터리 식별 번호
	Status : UDINT; // 배터리 전체 상태 비트
	OnlineRackCount : UDINT; // 통신 정상으로 판단한 랙 수
	TotalRackCount : UDINT; // 설치된 전체 랙 수
	MaxCellVoltageLocationFromRack : UDINT; // 최대 셀 전압 발생 위치의 랙 번호
	MaxCellVoltageLocationFromModule : UDINT; // 최대 셀 전압 발생 위치의 모듈 번호
	MaxCellVoltageLocationFromCell : UDINT; // 최대 셀 전압 발생 위치의 셀 번호
	MinCellVoltageLocationFromRack : UDINT; // 최소 셀 전압 발생 위치의 랙 번호
	MinCellVoltageLocationFromModule : UDINT; // 최소 셀 전압 발생 위치의 모듈 번호
	MinCellVoltageLocationFromCell : UDINT; // 최소 셀 전압 발생 위치의 셀 번호
	MaxModuleTempLocationFromRack : UDINT; // 모듈 최고 온도 발생 위치의 랙 번호
	MaxModuleTempLocationFromModule : UDINT; // 모듈 최고 온도 발생 위치의 모듈 번호
	MaxModuleTempLocationFromCell : UDINT; // 모듈 최고 온도 발생 위치의 셀 번호
	MinModuleTempLocationFromRack : UDINT; // 모듈 최저 온도 발생 위치의 랙 번호
	MinModuleTempLocationFromModule : UDINT; // 모듈 최저 온도 발생 위치의 모듈 번호
	MinModuleTempLocationFromCell : UDINT; // 모듈 최저 온도 발생 위치의 셀 번호
	Heartbeat : UDINT; // BMS 데이터 갱신 카운터
	Soc : REAL; // 배터리 충전 상태
	Soh : REAL; // 배터리 건강 상태
	Eol : REAL; // 배터리 수명 종료 관련 값
	DcVoltage : REAL; // 배터리 전체 직류 전압
	DcCurrent : REAL; // 배터리 전체 직류 전류
	ChargeCurrentLimit : REAL; // 배터리 전체 충전 허용 전류
	DischargeCurrentLimit : REAL; // 배터리 전체 방전 허용 전류
	ChargePowerLimit : REAL; // 배터리 전체 충전 허용 전력
	DischargePowerLimit : REAL; // 배터리 전체 방전 허용 전력
	MaxCellVoltage : REAL; // 전체 셀 중 최대 전압
	MinCellVoltage : REAL; // 전체 셀 중 최소 전압
	MaxModuleTemperature : REAL; // 전체 모듈 중 최고 온도
	MinModuleTemperature : REAL; // 전체 모듈 중 최저 온도
	Warning1 : UDINT; // 배터리 경보 비트 묶음 1
	Warning2 : UDINT; // 배터리 경보 비트 묶음 2
	Warning3 : UDINT; // 배터리 경보 비트 묶음 3
	Warning4 : UDINT; // 배터리 경보 비트 묶음 4
	Warning5 : UDINT; // 배터리 경보 비트 묶음 5
	Warning6 : UDINT; // 배터리 경보 비트 묶음 6
	Warning7 : UDINT; // 배터리 경보 비트 묶음 7
	Warning8 : UDINT; // 배터리 경보 비트 묶음 8
	Warning9 : UDINT; // 배터리 경보 비트 묶음 9
	Warning10 : UDINT; // 배터리 경보 비트 묶음 10
	Fault1 : UDINT; // 배터리 고장 비트 묶음 1
	Fault2 : UDINT; // 배터리 고장 비트 묶음 2
	Fault3 : UDINT; // 배터리 고장 비트 묶음 3
	Fault4 : UDINT; // 배터리 고장 비트 묶음 4
	Fault5 : UDINT; // 배터리 고장 비트 묶음 5
	Fault6 : UDINT; // 배터리 고장 비트 묶음 6
	Fault7 : UDINT; // 배터리 고장 비트 묶음 7
	Fault8 : UDINT; // 배터리 고장 비트 묶음 8
	Fault9 : UDINT; // 배터리 고장 비트 묶음 9
	Fault10 : UDINT; // 배터리 고장 비트 묶음 10
END_STRUCT
END_TYPE

// ---- 20_Module/Mqtt/Publish/ST_EssPublish_V1.TcDUT
{attribute 'pack_mode' := '1'}
TYPE ST_EssPublish_V1 :
STRUCT
	DeviceIndex	:	UDINT;
	Status	:	UDINT;
	AcActivePower	:	REAL;
	AcReactivePower:	REAL;
	AcVoltageR     :	REAL;
	AcVoltageS     :	REAL;
	AcVoltageT     :	REAL;
	AcCurrentR     :	REAL;
	AcCurrentS     :	REAL;
	AcCurrentT     :	REAL;
	Frequency      :	REAL;
	PowerFactor    :	REAL;
	EnergyActivePower:	REAL;
	EnergyReactivePower:	REAL;
	EnergyReverseActivePower:	REAL;
	EnergyReverseReactivePower:	REAL;
	Warning1:	UDINT;
	Warning2:	UDINT;
	Warning3:	UDINT;
	Warning4:	UDINT;
	Warning5:	UDINT;
	Warning6:	UDINT;
	Warning7:	UDINT;
	Warning8:	UDINT;
	Warning9:	UDINT;
	Warning10:	UDINT;
	Fault1:		UDINT;
	Fault2:		UDINT;
	Fault3:		UDINT;
	Fault4:		UDINT;
	Fault5:		UDINT;
	Fault6:		UDINT;
	Fault7:		UDINT;
	Fault8:		UDINT;
	Fault9:		UDINT;
	Fault10:		UDINT;
END_STRUCT
END_TYPE

// ---- 20_Module/Mqtt/Publish/ST_PcsPublish_V1.TcDUT
{attribute 'pack_mode' := '1'}
TYPE ST_PcsPublish_V1 :
STRUCT
	DeviceIndex			:	UDINT;
	SystemOperationMode	:	UDINT;	// 0: 수동, 1: 모드스케줄
	OperationMode			:	UDINT;
	PMSActivePower			:	REAL;	// kW
	RemoteMode				:	UDINT;	// 0: Local, 1: Remote
	Status					:	UDINT;	// bit0~9
	AcActivePower			:	REAL;	// kW
	AcReactivePower			:	REAL;	// kVar
	PowerFactor				:	REAL;
	Frequency				:	REAL;	// Hz
	AcRsVoltage				:	REAL;	// V
	AcStVoltage				:	REAL;	// V
	AcTrVoltage				:	REAL;	// V
	AcRVoltage				:	REAL;	// V
	AcSVoltage				:	REAL;	// V
	AcTVoltage				:	REAL;	// V
	AcRCurrent				:	REAL;	// A
	AcSCurrent				:	REAL;	// A
	AcTCurrent				:	REAL;	// A
	DcLinkVoltage			:	REAL;	// V
	DcVoltage				:	REAL;	// V
	DcCurrent				:	REAL;	// A
	DcActivePower			:	REAL;	// kW
	InsulationResistance	:	REAL;	// kΩ
	Temperature1			:	REAL;
	Temperature2			:	REAL;
	Temperature3			:	REAL;
	Temperature4			:	REAL;
	Temperature5			:	REAL;
	Temperature6			:	REAL;
	Temperature7			:	REAL;
	Temperature8			:	REAL;
	Warning1				:	UDINT;
	Warning2				:	UDINT;
	Warning3				:	UDINT;
	Warning4				:	UDINT;
	Warning5				:	UDINT;
	Warning6				:	UDINT;
	Warning7				:	UDINT;
	Warning8				:	UDINT;
	Warning9				:	UDINT;
	Warning10				:	UDINT;
	Fault1					:	UDINT;
	Fault2					:	UDINT;
	Fault3					:	UDINT;
	Fault4					:	UDINT;
	Fault5					:	UDINT;
	Fault6					:	UDINT;
	Fault7					:	UDINT;
	Fault8					:	UDINT;
	Fault9					:	UDINT;
	Fault10					:	UDINT;
END_STRUCT
END_TYPE

// ---- 20_Module/Mqtt/Publish/ST_PmsPublish_V1.TcDUT
{attribute 'pack_mode' := '1'}
TYPE ST_PmsPublish_V1 :
STRUCT
	DeviceIndex			:	UDINT;
	Status				:	UDINT;
	PmsIsAlive			:	UDINT;		// 0: 비정상, 1: 정상
	CpuUsage			:	UDINT;		// %
	CpuTemperature		:	UDINT;		// ℃
	RemainCycle			:	UDINT;		// %
	RemainSaveArea		:	UDINT;		// %
	ProtectModuleCurrent:	REAL;
	ProtectModuleVoltage:	REAL;
	PmsEvent			:	UDINT;
	ModuleStatus1		:	UDINT;
	ModuleStatus2		:	UDINT;
END_STRUCT
END_TYPE

// ---- 20_Module/Mqtt/Publish/ST_PvPublish_V1.TcDUT
{attribute 'pack_mode' := '1'}
TYPE ST_PvPublish_V1 :
STRUCT
	DeviceIndex	:	UDINT;
	Status		:	UDINT;
	AcActivePower						:			REAL;
	AcReactivePower                     :		    real;
	AcVoltageR                          :		    real;
	AcVoltageS                          :		    real;
	AcVoltageT                          :		    real;
	AcCurrentR                          :		    real;
	AcCurrentS                          :		    real;
	AcCurrentT                          :		    real;
	Frequency                           :		    real;
	PowerFactor                         :		    real;
	EnergyActivePower                   :		    real;
	EnergyReactivePower                 :		    real;
	EnergyReverseActivePower            :		    real;
	EnergyReverseReactivePower          :		    real;
	Warning1                            :			UDINT;
	Warning2                            :			UDINT;
	Warning3                            :			UDINT;
	Warning4                            :			UDINT;
	Warning5                            :			UDINT;
	Warning6                            :			UDINT;
	Warning7                            :			UDINT;
	Warning8                            :			UDINT;
	Warning9                            :			UDINT;
	Warning10                           :			UDINT;
	Fault1                              :			UDINT;
	Fault2                              :			UDINT;
	Fault3                              :			UDINT;
	Fault4                              :			UDINT;
	Fault5                              :			UDINT;
	Fault6                              :			UDINT;
	Fault7                              :			UDINT;
	Fault8                              :			UDINT;
	Fault9                              :			UDINT;
	Fault10                             :			UDINT;
END_STRUCT
END_TYPE

// ---- 20_Module/Mqtt/Publish/ST_RackPublish_V1.TcDUT
{attribute 'pack_mode' := '1'}
TYPE ST_RackPublish_V1 :
STRUCT
	DeviceIndex : UDINT;
	BatIndex : UDINT;
	Status : UDINT;
	ModuleCount : UDINT;
	Soc : REAL;
	Soh : REAL;
	DcVoltage : REAL;
	DcCurrent : REAL;
	ChargeCurrentLimit : REAL;
	DischargeCurrentLimit : REAL;
	ChargePowerLimit : REAL;
	DischargePowerLimit : REAL;
	AvgCellVoltage : REAL;
	MaxCellVoltage : REAL;
	MinCellVoltage : REAL;
	AvgModuleTemp : REAL;
	MaxModuleTemp : REAL;
	MinModuleTemp : REAL;
	MaxCellVoltageLocationFromModule : UDINT;
	MaxCellVoltageLocationFromCell : UDINT;
	MinCellVoltageLocationFromModule : UDINT;
	MinCellVoltageLocationFromCell : UDINT;
	MaxModuleTempLocationFromModule : UDINT;
	MaxModuleTempLocationFromCell : UDINT;
	MinModuleTempLocationFromModule : UDINT;
	MinModuleTempLocationFromCell : UDINT;
	Warning1 : UDINT;
	Warning2 : UDINT;
	Warning3 : UDINT;
	Warning4 : UDINT;
	Warning5 : UDINT;
	Warning6 : UDINT;
	Warning7 : UDINT;
	Warning8 : UDINT;
	Warning9 : UDINT;
	Warning10 : UDINT;
	Fault1 : UDINT;
	Fault2 : UDINT;
	Fault3 : UDINT;
	Fault4 : UDINT;
	Fault5 : UDINT;
	Fault6 : UDINT;
	Fault7 : UDINT;
	Fault8 : UDINT;
	Fault9 : UDINT;
	Fault10 : UDINT;
END_STRUCT
END_TYPE

// ---- 20_Module/Mqtt/Publish/ST_TempPublish_V1.TcDUT
{attribute 'pack_mode' := '1'}
TYPE ST_TempPublish_V1 :
STRUCT
	DeviceIndex	:	UDINT;
	status		:	UDINT;
	location	:	UDINT;		//1: PCS 실 2: BAT 실 3: UPS 실 4: FC 컨테이너 실 5: 외부
	temperature	:	REAL;
	humidity	:	REAL;
END_STRUCT
END_TYPE

// ---- 20_Module/Mqtt/Publish/ST_AirConditionerPublishData.TcDUT
{attribute 'pack_mode' := '1'}
TYPE ST_AirConditionerPublishData :
STRUCT
	Header		:	ST_MqttHeader;
	Devices		:	ARRAY[0..GVL_PARAM.AIR_CONDITIONER_COUNT-1] OF ST_AirConditionerPublish_V1;
END_STRUCT
END_TYPE

// ---- 20_Module/Mqtt/Publish/ST_BatPublishData.TcDUT
{attribute 'pack_mode' := '1'}
TYPE ST_BatPublishData :
STRUCT
	Header		:	ST_MqttHeader;
	Devices		:	ARRAY[0..GVL_PARAM.BMS_COUNT-1] OF ST_BatPublish_V1;
END_STRUCT
END_TYPE

// ---- 20_Module/Mqtt/Publish/ST_EssPublishData.TcDUT
{attribute 'pack_mode' := '1'}
TYPE ST_EssPublishData :
STRUCT
	Header		:	ST_MqttHeader;
	Devices		:	ARRAY[0..GVL_PARAM.ESS_COUNT-1] OF ST_EssPublish_V1;
END_STRUCT
END_TYPE

// ---- 20_Module/Mqtt/Publish/ST_PcsPublishData.TcDUT
{attribute 'pack_mode' := '1'}
TYPE ST_PcsPublishData :
STRUCT
	Header		:	ST_MqttHeader;
	Devices		:	ARRAY[0..GVL_PARAM.PCS_COUNT-1] OF ST_PcsPublish_V1;
END_STRUCT
END_TYPE

// ---- 20_Module/Mqtt/Publish/ST_PmsPublishData.TcDUT
{attribute 'pack_mode' := '1'}
TYPE ST_PmsPublishData :
STRUCT
	Header		:	ST_MqttHeader;
	Devices		:	ARRAY[0..0] OF ST_PmsPublish_V1;
END_STRUCT
END_TYPE

// ---- 20_Module/Mqtt/Publish/ST_PvPublishData.TcDUT
{attribute 'pack_mode' := '1'}
TYPE ST_PvPublishData :
STRUCT
	Header		:	ST_MqttHeader;
	Devices		:	ARRAY[0..GVL_PARAM.PV_COUNT-1] OF ST_PvPublish_V1;
END_STRUCT
END_TYPE

// ---- 20_Module/Mqtt/Publish/ST_RackPublishData.TcDUT
{attribute 'pack_mode' := '1'}
TYPE ST_RackPublishData :
STRUCT
	Header		:	ST_MqttHeader;
	Devices		:	ARRAY[0..GVL_PARAM.RACK_COUNT-1] OF ST_RackPublish_V1;
END_STRUCT
END_TYPE

// ---- 20_Module/Mqtt/Publish/ST_TempPublishData.TcDUT
{attribute 'pack_mode' := '1'}
TYPE ST_TempPublishData :
STRUCT
	Header		:	ST_MqttHeader;
	Devices		:	ARRAY[0..GVL_PARAM.TEMP_COUNT-1] OF ST_TempPublish_V1;
END_STRUCT
END_TYPE

// ---- 20_Module/Mqtt/Config/ST_BatConfig_Rx.TcDUT
{attribute 'pack_mode' := '1'}
TYPE ST_BatConfig_Rx :
STRUCT
	DeviceId : UDINT;
	SocMin : REAL;
	SocMax : REAL;
END_STRUCT
END_TYPE

// ---- 20_Module/Mqtt/Config/ST_CommonConfig_REAL.TcDUT
TYPE ST_CommonConfig_REAL :
STRUCT
	value	: REAL;
	is_available : UDINT;
END_STRUCT
END_TYPE

// ---- 20_Module/Mqtt/Config/ST_CommonConfig_UDINT.TcDUT
TYPE ST_CommonConfig_UDINT :
STRUCT
	value	: UDINT;
	is_available : UDINT;
END_STRUCT
END_TYPE

// ---- 20_Module/Mqtt/Config/ST_PcsConfig_Rx.TcDUT
{attribute 'pack_mode' := '1'}
TYPE ST_PcsConfig_Rx :
STRUCT
	DeviceId			:	UDINT;
	ChargePowerLimit	:	ST_CommonConfig_UDINT;	// kW
	DisChargePowerLimit	:	ST_CommonConfig_UDINT;	// kW
	PvMarginRate		:	ST_CommonConfig_UDINT;	// %
END_STRUCT
END_TYPE

// ---- 20_Module/Mqtt/Config/ST_ProtectionConfig_Rx.TcDUT
{attribute 'pack_mode' := '1'}
TYPE ST_ProtectionConfig_Rx :
STRUCT
	BatWarrning			:	REAL;
	BatFault			:	REAL;
	BatRoomTempWarrning	:	REAL;
	BatRoomTempFault	:	REAL;
	BatRoomHumWarrning	:	REAL;
	BatRoomHumFault		:	REAL;
END_STRUCT
END_TYPE

// ---- 20_Module/Mqtt/Config/ST_BatConfigWirePacket.TcDUT
{attribute 'pack_mode' := '1'}
TYPE ST_BatConfigWirePacket :
STRUCT
	Header	:	ST_MqttCommandHeader;
	Records	:	ARRAY[0..GVL_PARAM.BMS_COUNT-1] OF ST_BatConfig_Rx;
END_STRUCT
END_TYPE

// ---- 20_Module/Mqtt/Config/ST_PcsConfigWirePacket.TcDUT
{attribute 'pack_mode' := '1'}
TYPE ST_PcsConfigWirePacket :
STRUCT
	Header	:	ST_MqttCommandHeader;
	Records	:	ARRAY[0..GVL_PARAM.PCS_COUNT-1] OF ST_PcsConfig_Rx;
END_STRUCT
END_TYPE

// ---- 20_Module/Mqtt/Config/ST_ProtectionConfigWirePacket.TcDUT
{attribute 'pack_mode' := '1'}
TYPE ST_ProtectionConfigWirePacket :
STRUCT
	Header	:	ST_MqttCommandHeader;
	Record	:	ST_ProtectionConfig_Rx;	// DeviceIndex 없는 단일 레코드
END_STRUCT
END_TYPE

// ---- 20_Module/Mqtt/ST_IfEmsCmd.TcDUT
TYPE ST_IfEmsCmd :		// MQTT → MAIN 명령 칸 (GVL_IF.g_stEmsCmd). 쓰는 곳: PRG_Mqtt (FB_EmsCommand 결과), 읽는 곳: FB_SrcEms
STRUCT
	nRxCount		: UDINT;		// 받은 command 메시지 누계 (브로커 3개 합). 명령이 없는 메시지도 셈 → EMS가 살아 있다는 표시
	astPcs			: ARRAY[1..GVL_PARAM.PCS_COUNT] OF ST_PcsCmd;	// PCS 상태 명령 + 번호 (칸 = PCS 번호 = DeviceIndex + 1)
	afPcsP			: ARRAY[1..GVL_PARAM.PCS_COUNT] OF REAL;		// 충전·방전 P 지령 kW (방전 +, 충전 −). PCS 한 대 몫
	anPcsPSeq		: ARRAY[1..GVL_PARAM.PCS_COUNT] OF UDINT;		// P 지령 번호. 바뀌면 새 지령 (0 = 한 번도 못 받음)
	astBatRack		: ARRAY[1..GVL_PARAM.BMS_COUNT] OF ST_BatRackCmd;	// 랙 컨택터 명령 (CommandType 11·12). MAIN → FB_BmsRackCommand
	astBatCtl		: ARRAY[1..GVL_PARAM.BMS_COUNT] OF ST_BatCtlCmd;	// 컨택터 하나씩 명령 (CommandType 5~10). MAIN → FB_BmsContactorCommand [2026-11-13]
	astBat			: ARRAY[1..GVL_PARAM.BMS_COUNT] OF ST_BatCmd;	// BMS 명령 + 번호 (칸 = BMS 번호 = DeviceIndex + 1)
END_STRUCT
END_TYPE

// ---- 20_Module/Mqtt/ST_MqttBroker.TcDUT
TYPE ST_MqttBroker :		// 브로커 한 곳의 접속 설정
STRUCT
	bUse		: BOOL;				// FALSE = 이 브로커에 접속하지 않음
	sHost		: STRING(15);		// IP 주소
	nPort		: UINT := 1883;
END_STRUCT
END_TYPE

// ---- 20_Module/Mqtt/ST_MqttSet.TcDUT
TYPE ST_MqttSet :		// MQTT 접속 설정 (현장마다 다름. GVL_SITE.MQTT_SET → FB_MqttMain.i_stSet)
STRUCT
	nSiteId			: UDINT;			// 사이트 번호 (토픽·헤더·ClientId에 들어감)
	stCloud			: ST_MqttBroker;
	stLocal			: ST_MqttBroker;
	stAzure			: ST_MqttBroker;
	sUserName		: STRING;			// 브로커 계정 (세 브로커 공통)
	sUserPassword	: STRING;
END_STRUCT
END_TYPE

// ---- 20_Module/Mqtt/ST_IfReport.TcDUT
TYPE ST_IfReport :		// MAIN → MQTT 보고 칸 (GVL_IF.g_stReport). 쓰는 곳: MAIN 액션 A_Report (PCS·BAT 보고 매핑 결과), 읽는 곳: PRG_Mqtt
STRUCT
	abPcsMapped		: ARRAY[1..GVL_PARAM.PCS_COUNT] OF BOOL;			// 이 PCS를 매핑 모듈이 채움. FALSE면 PRG_Mqtt는 발행 구조체를 건드리지 않음 (시험 더미 유지)
	abPcsComm		: ARRAY[1..GVL_PARAM.PCS_COUNT] OF BOOL;			// 통신 정상. FALSE면 astPcs는 모두 0
	astPcs			: ARRAY[1..GVL_PARAM.PCS_COUNT] OF ST_PcsPublish_V1;	// 발행 직전 레코드 (칸 = PCS 번호 = 발행 DeviceIndex, 1부터)
	abBatMapped : ARRAY[1..GVL_PARAM.BMS_COUNT] OF BOOL; // BAT 매핑 연결 여부
	abBatValid : ARRAY[1..GVL_PARAM.BMS_COUNT] OF BOOL; // BAT 데이터 유효 여부
	astBat : ARRAY[1..GVL_PARAM.BMS_COUNT] OF ST_BatPublish_V1; // BAT 보고값
	astRack : ARRAY[1..GVL_PARAM.RACK_COUNT] OF ST_RackPublish_V1; // RACK 보고값. abBatMapped를 따름
	astModule : ARRAY[1..GVL_PARAM.BAT_MODULE_COUNT] OF ST_ModulePublish_V1; // MODULE 보고값. abBatMapped를 따름
	abUpsMapped : ARRAY[1..GVL_PARAM.UPS_COUNT] OF BOOL; // UPS 매핑 연결 여부
	abUpsValid : ARRAY[1..GVL_PARAM.UPS_COUNT] OF BOOL; // UPS 데이터 유효 여부
	astUps : ARRAY[1..GVL_PARAM.UPS_COUNT] OF ST_UpsPublish_V1; // UPS 보고값
	abImdMapped : ARRAY[1..GVL_PARAM.IMD_COUNT] OF BOOL; // IMD 매핑 연결 여부
	abImdValid : ARRAY[1..GVL_PARAM.IMD_COUNT] OF BOOL; // IMD 데이터 유효 여부
	astImd : ARRAY[1..GVL_PARAM.IMD_COUNT] OF ST_ImdPublish_V1; // IMD 보고값
	abFireMapped : ARRAY[1..GVL_PARAM.FIRE_COUNT] OF BOOL; // 화재감지기 매핑 연결 여부
	astFire : ARRAY[1..GVL_PARAM.FIRE_COUNT] OF ST_FirePublish_V1; // 화재감지기 보고값
	abTempMapped : ARRAY[1..GVL_PARAM.TEMP_COUNT] OF BOOL; // 온습도 매핑 연결 여부
	astTemp : ARRAY[1..GVL_PARAM.TEMP_COUNT] OF ST_TempPublish_V1; // 온습도 보고값
END_STRUCT
END_TYPE

// ---- 20_Module/Mqtt/Logger/ST_LoggerHeader.TcDUT
{attribute 'pack_mode' := '1'}
TYPE ST_LoggerHeader :		// 로거 토픽(pms_log) 헤더 (36 byte). 장치 토픽 헤더(ST_MqttHeader)와 달리 DeviceCount 없음: 메시지 1건 = 이벤트 1건
STRUCT
	HeaderVersion	:	UDINT;		// GVL_MQTT.HEADER_VERSION
	DeviceVersion	:	UDINT;		// GVL_MQTT.LOGGER_VERSION
	SiteId			:	UDINT;
	TimeStamp		:	STRING(23);	// 이벤트가 생긴 시각 (보낸 시각 아님, 현지 시각) "2024-09-04 11:11:11.123" (23자 + null = 24byte)
END_STRUCT
END_TYPE

// ---- 20_Module/Mqtt/Logger/ST_LoggerPublish_V1.TcDUT
{attribute 'pack_mode' := '1'}
TYPE ST_LoggerPublish_V1 :		// 로거 토픽 패킷 (238 byte): 헤더 + 로그 문구. dgspms/{solution}/{사이트}/{LOGGER_TOPIC} (지금 pms_log)
STRUCT
	Header		:	ST_LoggerHeader;	// 36 byte
	Contents	:	WSTRING(100);		// 로그 문구 (UTF-16LE, 100자 + null = 202 byte). 알람 해소는 앞에 '[해소] '. 길이는 GVL_MQTT.LOGGER_TEXT_MAX와 같게
END_STRUCT
END_TYPE

// ---- 20_Module/Mqtt/Logger/ST_LoggerSlot.TcDUT
TYPE ST_LoggerSlot :		// 로거 큐 한 칸 (FB_MqttLoggerListener 안에서만 씀)
STRUCT
	nNo				: UDINT;		// 이벤트 번호 (받은 순서, 1부터). 0 = 빈 칸
	nTimestamp		: ULINT;		// 로거 기록 시각 (FILETIME: UTC, 100 ns)
	nEventId		: UDINT;		// 이벤트 ID (문구를 못 받았을 때 대체 문구에 씀)
	bCleared		: BOOL;			// 알람 해소
	bRequesting		: BOOL;			// 문구 요청 중 (같은 칸 번호의 FB_RequestEventText)
	nRequestStart	: ULINT;		// 문구 요청 시작 (F_GetSystemTime). 너무 오래 걸리면 대체 문구
	bTextDone		: BOOL;			// 문구 받음
	bReady			: BOOL;			// 발행 준비 끝 (문구 + 시각 문자열)
	sTime			: STRING(23);	// 현지 시각 문자열
	wsText			: WSTRING(100);	// 발행할 문구 (해소 표시 포함, 100자 이내)
END_STRUCT
END_TYPE

// ---- 10_Core/00_Type/E_CtrlModeRefuse.TcDUT
{attribute 'strict'}
TYPE E_CtrlModeRefuse :		// 제어 모드 요청 결과
(
	None		:= 0,	// 접수 (또는 이미 켜져 있음)
	BadSlot		:= 1,	// 칸 번호가 범위 밖이거나 빈 칸
	NotReady	:= 2	// 모드의 진입 조건이 안 맞음 (이유 코드 q_nRefuseReason → 그 모드의 M_ReasonText)
) INT;
END_TYPE

// ---- 10_Core/00_Type/E_CtrlModeStep.TcDUT
{attribute 'strict'}
TYPE E_CtrlModeStep :		// 제어 모드 관리자 단계
(
	Idle		:= 0,	// 켜진 모드 없음 (지령을 내지 않음)
	Active		:= 1,	// 모드 하나가 동작 중
	Leaving		:= 2	// 전환 중: 이전 모드는 끝났고 그 모드가 내던 P·Q를 0으로 둠 (ST_CtrlModeSet.tZeroDelay)
) INT;
END_TYPE

// ---- 10_Core/00_Type/ST_CtrlModeOut.TcDUT
TYPE ST_CtrlModeOut :		// 제어 모드 한 스캔 결과 (I_ControlMode.M_Calc)
STRUCT
	bPSetActive	: BOOL;
	fPSet		: REAL;			// kW, 접속점 기준 (방전 +)
	bQSetActive	: BOOL;
	fQSet		: REAL;			// kvar, 접속점 기준 (공급 +)
	bExitReq	: BOOL;			// 모드가 스스로 끝냄 (운전 시간 끝, 필요한 계측 무효 등). 관리자가 M_Exit를 부르고 대체 모드로 넘어감
	nReason		: UINT;			// 끝낸 이유 코드 (그 모드의 M_ReasonText)
	(* [16번 수정 2026-11-09: 추가] 유닛별 값. 접속점 그룹 단위 관리자에서 PCS마다 다른 값을 내는 모드(스탠다드 스케줄: EMS가 PCS마다 지령)가 씀 *)
	bUnitOut	: BOOL;			// TRUE = astUnit을 냄 (접속점 그룹 값 bPSetActive·fPSet·bQSetActive·fQSet은 쓰지 않음)
	astUnit		: ARRAY[1..GVL_PARAM.UNIT_COUNT] OF ST_UnitReq;	// 유닛 출력 (kW·kvar). 접속점 그룹 단위 관리자는 전부, 유닛 단위 관리자는 맡은 유닛 칸만 냄
END_STRUCT
END_TYPE

// ---- 10_Core/00_Type/ST_CtrlModeSet.TcDUT
TYPE ST_CtrlModeSet :		// 제어 모드 관리자 설정 (GVL_PERSIST.g_stModuleSet 칸 → A_PassModuleSet)
STRUCT
	bZeroOnSwitch	: BOOL := TRUE;		// 모드를 바꿀 때 이전 모드가 내던 P·Q를 0으로 둔 뒤 새 모드 진입. FALSE = 바로 진입 (출력 변화는 그룹 램프 bRamp가 맡음)
	tZeroDelay		: TIME := T#1S;		// 0으로 두는 시간
	nFallback		: UINT;				// 켜진 모드가 스스로 끝낼 때 넘어갈 칸 번호. 0 = 모드 없음
	ePccShare		: E_PccShare := E_PccShare.ByRating;	// 유닛 단위(FB_CtrlModeMgr.i_nUnit ≠ 0)일 때 모드가 보는 접속점 값 (그룹 단위에서는 안 씀)
	fPccRatio		: REAL := 1.0;		// ePccShare = Fixed일 때 이 유닛 몫 (0~1)
END_STRUCT
END_TYPE

// ---- 20_Module/ControlMode/ST_CmConstPowerSet.TcDUT
TYPE ST_CmConstPowerSet :	// 정출력 모드 설정
STRUCT
	fPSet		: REAL;			// kW, 접속점 기준 (방전 +, 충전 -)
	bQSet		: BOOL;			// Q도 냄 (FALSE = Q는 다른 지령원에 맡김)
	fQSet		: REAL;			// kvar, 접속점 기준 (공급 +)
	tDuration	: TIME;			// 운전 시간. T#0S = 끝없이 (요청이 바뀔 때까지)
END_STRUCT
END_TYPE

// ---- 20_Module/ControlMode/ST_CmExtCmd.TcDUT
TYPE ST_CmExtCmd :		// 바깥(EMS 등)에서 받은 지령 한 대 몫 (FB_CmStdSchedule 입력). MAIN이 지령원 결과에서 채움 (이 모드는 통신 형식을 모름)
STRUCT
	bUse		: BOOL;			// 이 칸(유닛)에 지령을 냄 (이 모드가 맡은 유닛). [16번 수정 2026-11-09: 추가 — 모드가 유닛마다 칸을 받음]
	bAlive		: BOOL;			// 바깥 지령원이 살아 있음 (끊기면 받아 둔 P를 버리고 0)
	nPSeq		: UDINT;		// P 지령 번호. 바뀌면 새 P 지령
	fP			: REAL;			// kW, P 지령 (방전 +, 충전 -). 이 유닛 출력
	nStateSeq	: UDINT;		// 상태 명령 번호. 바뀌면 새 상태 명령
	eState		: E_PcsCmd;		// 마지막 상태 명령 (Stop·Standby·EStop이면 받아 둔 P를 버림)
END_STRUCT
END_TYPE

// ---- 10_Core/00_Type/ST_LocalTime.TcDUT
TYPE ST_LocalTime :		// 현지 시각 (플랫폼과 무관한 모양. TwinCAT은 20_Module\Common\FB_LocalClock이 채움)
STRUCT
	bValid		: BOOL;		// 시각을 믿을 수 있음 (첫 동기 뒤). FALSE면 아래 값을 쓰지 않음
	nYear		: UINT;
	nMonth		: UINT;		// 1~12
	nDay		: UINT;		// 1~31
	nDayOfWeek	: UINT;		// 0 = 일요일 ~ 6 = 토요일
	nHour		: UINT;		// 0~23
	nMinute		: UINT;		// 0~59
	nSecond		: UINT;		// 0~59
END_STRUCT
END_TYPE

// ---- 10_Core/00_Type/ST_CtrlModeView.TcDUT
TYPE ST_CtrlModeView :		// 제어 모드에 넘기는 값 (FB_CtrlModeMgr가 매 스캔 채움). 필요한 값이 늘면 칸을 더함 (모드는 고치지 않아도 됨)
STRUCT
	stGroup		: ST_GroupView;		// 대상 그룹 값 (접속점 계측·정격·가용·SOC·실제 출력)
	stTime		: ST_LocalTime;		// 현지 시각
END_STRUCT
END_TYPE

// ---- 20_Module/Mqtt/E_MqttBroker.TcDUT
{attribute 'qualified_only'}
{attribute 'strict'}
TYPE E_MqttBroker :		// MQTT 브로커 (GVL_SITE.MQTT_SET의 stCloud·stLocal·stAzure) [9번 수정 2026-11-09: 추가]
(
	Cloud	:= 1,
	Local	:= 2,
	Azure	:= 3
) INT;
END_TYPE

// ---- 20_Module/Mqtt/ST_BrokerWatchSet.TcDUT
TYPE ST_BrokerWatchSet :		// MQTT 브로커 끊김 감시 설정 (GVL_PERSIST.g_stBrokerWatch, 운전 중 바꿈·이중화 동기화) [9번 수정 2026-11-09: 추가]
STRUCT
	eBroker		: E_MqttBroker := E_MqttBroker.Local;	// 감시할 브로커. MQTT_SET에서 쓰지 않는(bUse FALSE) 브로커를 고르면 감시하지 않음
	tLostDelay	: TIME := T#30S;		// 접속이 이 시간 넘게 끊기면 '브로커 끊김' 알람 + 운전 모드 요청을 모두 Manual로 (끊김마다 한 번)
END_STRUCT
END_TYPE

// ---- 20_Module/Mqtt/ST_IfEmsCfg.TcDUT
TYPE ST_IfEmsCfg :		// MQTT → MAIN config 칸 (GVL_IF.g_stEmsCfg). 쓰는 곳: PRG_Mqtt, 읽는 곳: FB_EmsConfigApply [9-21 수정 2026-11-04: 추가]
STRUCT
	astPcs		: ARRAY[1..GVL_PARAM.PCS_COUNT] OF ST_PcsConfig_Rx;	// 마지막으로 받은 config/pcs 레코드 (칸 = PCS 번호 = DeviceId + 1)
	anPcsSeq	: ARRAY[1..GVL_PARAM.PCS_COUNT] OF UDINT;			// 그 칸에 새 레코드가 들어올 때마다 1 올림 (0 = 한 번도 못 받음)
	astBat		: ARRAY[1..GVL_PARAM.BMS_COUNT] OF ST_BatConfig_Rx;	// 마지막으로 받은 config/bat 레코드 (칸 = BMS 번호 = DeviceId + 1)
	anBatSeq	: ARRAY[1..GVL_PARAM.BMS_COUNT] OF UDINT;
END_STRUCT
END_TYPE

// ---- 20_Module/Mqtt/ST_IfEmsCfgEcho.TcDUT
TYPE ST_IfEmsCfgEcho :		// MAIN → MQTT config echo 칸 (GVL_IF.g_stEmsCfgEcho). 실제 설정을 config 레코드 모양으로 (칸 = DeviceIndex). 쓰는 곳: MAIN (FB_EmsConfigApply.M_BuildEcho) [9-21 수정 2026-11-04: 추가]
STRUCT
	astPcs	: ARRAY[0..GVL_PARAM.PCS_COUNT-1] OF ST_PcsConfig_Rx;	// 충·방전 한도 = 그 PCS 유닛들의 사용자 한도 합 (모두 켜져 있으면 is_available 1). PvMarginRate = 받은 값, is_available 0 (PLC가 쓰지 않음)
	astBat	: ARRAY[0..GVL_PARAM.BMS_COUNT-1] OF ST_BatConfig_Rx;	// SOC 정책 상·하한 (버스 전체 한 세트라 BMS마다 같은 값)
END_STRUCT
END_TYPE

// ---- 20_Module/ControlMode/ST_SchedSlot.TcDUT
TYPE ST_SchedSlot :		// 시간표 한 칸
STRUCT
	nStart		: UINT;		// HHMM, 시작 (포함)
	nEnd		: UINT;		// HHMM, 끝 (미포함. 2400 = 자정까지). 시작 = 끝 = 빈 칸. 자정을 넘는 운전은 두 칸으로 (그날 ~2400, 다음날 0000~)
	fP			: REAL;		// kW, 접속점 기준 (방전 +, 충전 -). Messis 값(충전 +)과 부호가 반대
END_STRUCT
END_TYPE

// ---- 20_Module/ControlMode/ST_CmScheduleSet.TcDUT
TYPE ST_CmScheduleSet :		// 스케줄 시간표 (스케줄·통합 모드가 같은 표를 씀)
STRUCT
	astSlot		: ARRAY[0..2, 0..6, 1..GVL_PARAM.SCHED_SLOT_COUNT] OF ST_SchedSlot;	// [계절, 요일(0 = 일), 칸]. 맞는 칸이 여럿이면 번호가 큰 칸
END_STRUCT
END_TYPE

// ---- 10_Core/00_Type/E_PccShare.TcDUT
{attribute 'strict'}
TYPE E_PccShare :		// 유닛(PCS) 단위 제어 모드가 보는 접속점 값 (여러 유닛이 한 접속점을 같이 쓸 때. 유닛이 혼자인 그룹은 셋 다 같음)
(
	ByRating	:= 0,	// 그룹 부하(그룹 유닛 출력 합 - 접속점 P)를 가용 정격 비율로 나눈 몫만 봄. 몫 합 = 그룹 부하 → 피크컷·역송 방지가 겹치지 않음 (목표 피크도 몫으로 넣음)
	Actual		:= 1,	// 접속점 실측 그대로 (다른 유닛 출력이 들어간 값). 유닛마다 같은 수전을 보고 따로 반응 (피크컷이 겹칠 수 있음)
	Fixed		:= 2	// 정한 비율(ST_CtrlModeSet.fPccRatio, 0~1)로 나눈 몫
) INT;
END_TYPE

// ---- 10_Core/00_Type/ST_UnitView.TcDUT
TYPE ST_UnitView :		// 유닛(PCS) 하나 기준 값 (FB_UnitView). 유닛마다 둔 제어 모드 관리자(FB_CtrlModeMgr.i_nUnit ≠ 0)가 봄
STRUCT
	nUnit			: UINT;
	bAvail			: BOOL;				// 가용 (FB_UnitAvail)
	stView			: ST_GroupView;		// 유닛 기준. 정격·가용 한도·출력 = 이 유닛, 배터리 한도·용량 = 연결 버스 값을 버스 가용 유닛 정격 비율로 나눈 몫, SOC = 연결 배터리 그룹, 접속점(stPcc)·상태 = 소속 그룹 그대로
	fGroupPOut		: REAL;				// kW, 소속 그룹 유닛 출력 합 (실측). 접속점 몫 계산용 (그룹 부하 = 그룹 출력 - 접속점 P)
	fGroupQOut		: REAL;				// kvar
	fRatingShare	: REAL;				// 0~1, 소속 그룹 가용 P 한도 합 중 이 유닛 몫. 가용이 아니면 0
END_STRUCT
END_TYPE

// ---- 99_Test/ST_LoggerTestReg.TcDUT
TYPE ST_LoggerTestReg :		// PRG_TestLogger가 이벤트 로거에서 찾은 등록 이벤트 한 칸
STRUCT
	stEntry		: TcEventEntry;		// 클래스·번호 (심각도는 Info로 둠: 원래 심각도는 PLC에서 읽을 수 없음)
	wsName		: WSTRING(31);		// "클래스 번호" (예: PmsSystem 8)
	wsTemplate	: WSTRING(255);		// 받은 문구 틀 (인자 자리에 #0#~#5#)
	nArgs		: UINT;				// 인자 수
	nFixed		: UINT;				// 고정 글자 수 (인자를 뺀 길이)
	nFree		: INT;				// 95 − 고정 글자 = 인자에 쓸 수 있는 글자
	nPerArg		: UINT;				// 인자 하나당 남는 글자 (nFree / 인자 수)
	bCheck		: BOOL;				// 확인 필요: 고정 50자 초과 또는 인자 하나당 남는 글자 10자 미만
END_STRUCT
END_TYPE

// ---- 20_Module/ControlMode/ST_CmDisWindow.TcDUT
TYPE ST_CmDisWindow :		// 방전 허용 시간 (경부하 시간에는 방전하지 않음)
STRUCT
	bUse		: BOOL := TRUE;		// FALSE = 시간 제한 없음
	nStart		: UINT := 800;		// HHMM, 허용 시작 (포함)
	nEnd		: UINT := 2200;		// HHMM, 허용 끝 (미포함)
	bSunday		: BOOL := FALSE;	// 일요일 방전 허용 (기본: 일요일은 하루 종일 경부하)
END_STRUCT
END_TYPE

// ---- 20_Module/ControlMode/ST_CmNoReverse.TcDUT
TYPE ST_CmNoReverse :		// 역송 방지: 방전이 (부하 − 여유)를 넘으면 줄임. 부하 = ESS 출력(방전 +) − 접속점 공급
STRUCT
	bUse		: BOOL := TRUE;
	fMargin		: REAL := 10.0;		// kW, 남길 수전 여유 (Messis ReversePowerLimit + 10에 해당)
	fScale		: REAL := 0.95;		// 넘을 때 쓸 비율 (가능량 × 이 값)
END_STRUCT
END_TYPE

// ---- 20_Module/ControlMode/ST_CmCommonSet.TcDUT
TYPE ST_CmCommonSet :		// 요금제 기반 제어 모드 공통 설정 (스케줄·피크컷·통합이 같은 값을 씀)
STRUCT
	anSeasonOfMonth	: ARRAY[1..12] OF UINT := [2, 2, 1, 1, 1, 0, 0, 0, 1, 1, 2, 2];		// 월 → 계절 (0 여름, 1 봄·가을, 2 겨울). 기본 = 한전 계절
	abHoliday		: ARRAY[1..12, 1..31] OF BOOL;		// [월, 일] 휴일: 하루 종일 0
	stDis			: ST_CmDisWindow;	// 방전 허용 시간
	stNoRev			: ST_CmNoReverse;	// 역송 방지
END_STRUCT
END_TYPE

// ---- 20_Module/ControlMode/ST_CmPeakCalcSet.TcDUT
TYPE ST_CmPeakCalcSet :		// 15분 피크 제어 계산 (FB_CmPeakCalc)
STRUCT
	fTarget		: REAL;				// kW, 15분 평균 수전 목표 (계약·목표 피크). 0 = 피크 제어 안 함
	fBandSens	: REAL := 0.0;		// 시작 기준 감도: 부하가 목표 + 가용 출력 × (남은 분/15, 정수 나눗셈) × 이 값 × 0.5를 넘을 때만 제어. 0 = Messis 실제 동작 (목표를 넘으면 바로)
	fLoadRatio	: REAL := 0.8;		// 방전 상한 = 30초 평균 부하 × 이 값
	fMinOut		: REAL := 10.0;		// kW, 제어량이 1 kW를 넘으면 최소 이 값
END_STRUCT
END_TYPE

// ---- 20_Module/ControlMode/ST_CmWindowSet.TcDUT
TYPE ST_CmWindowSet :		// 시간 구간 + SOC (자동 충전: 채울 목표 SOC, 잔량 방전: 남길 하한 SOC)
STRUCT
	bUse		: BOOL;
	nStart		: UINT;		// HHMM (포함). 시작 > 끝이면 자정을 넘김
	nEnd		: UINT;		// HHMM (미포함). 이 시각까지 SOC를 맞추도록 출력을 정함
	fSoc		: REAL;		// %
END_STRUCT
END_TYPE

// ---- 20_Module/ControlMode/ST_CmPeakCutSet.TcDUT
TYPE ST_CmPeakCutSet :		// 피크컷 모드 설정
STRUCT
	stPeak		: ST_CmPeakCalcSet;
	stAutoChg	: ST_CmWindowSet := (fSoc := 100.0);	// 자동 충전 시간 (경부하 시간 충전). fSoc = 채울 목표
	stRemain	: ST_CmWindowSet := (fSoc := 10.0);		// 잔량 방전 시간 (남은 에너지를 끝 시각까지 고르게). fSoc = 남길 하한
END_STRUCT
END_TYPE

// ---- 20_Module/ControlMode/ST_CmSchedPeakSet.TcDUT
TYPE ST_CmSchedPeakSet :	// 통합 모드(스케줄 + 피크컷) 설정. 시간표는 스케줄 모드와 같은 표 (ST_CmScheduleSet)
STRUCT
	stPeak		: ST_CmPeakCalcSet;
	stRemain	: ST_CmWindowSet := (fSoc := 10.0);		// 잔량 방전 시간. fSoc = 남길 하한
END_STRUCT
END_TYPE

// ---- 20_Module/Driver/Plaspo/ST_PlaspoPcsRaw.TcDUT
TYPE ST_PlaspoPcsRaw :		// 플라스포 PCS 읽기 맵: 홀딩 레지스터 1번부터 39개 (Helios FB_PlaspoPcs와 같음)
STRUCT
	nPcsStatus		: WORD;		// 1: bit0 운전, bit1 고장, bit2 경고, bit5 PCS 내부 통신 이상
	nCdStatus		: UINT;		// 2: 0 대기, 1 충전, 2 방전
	nRemoteMode		: UINT;		// 3: 1 = 리모트 (PMS 제어 가능)
	nOpMode			: UINT;		// 4
	nRefFeedback	: UINT;		// 5
	nMmcStatus		: UINT;		// 6
	anFault			: ARRAY[1..5] OF WORD;		// 7~11 (5번째는 경고)
	anIgbtTemp		: ARRAY[1..4] OF INT;		// 12~15
	anAcFilterTemp	: ARRAY[1..4] OF INT;		// 16~19
	anAcVolt		: ARRAY[1..3] OF UINT;		// 20~22
	anAcCurrent		: ARRAY[1..3] OF UINT;		// 23~25
	nAcFreq			: UINT;		// 26: 0.1 Hz
	nAcActive		: INT;		// 27: 0.1 kW (Helios는 부호를 뒤집어 씀)
	nAcReactive		: INT;		// 28: 0.1 kvar
	nAcPf			: INT;		// 29
	nTodayDisEnergy	: UINT;		// 30
	nTodayChgEnergy	: UINT;		// 31
	nTotalDisH		: UINT;		// 32~35
	nTotalDisL		: UINT;
	nTotalChgH		: UINT;
	nTotalChgL		: UINT;
	nDcLinkVolt		: UINT;		// 36
	nDcVolt			: UINT;		// 37
	nDcCurrent		: INT;		// 38
	nDcPower		: INT;		// 39
END_STRUCT
END_TYPE

// ---- 10_Core/90_Redundancy/E_RedPeer.TcDUT
{attribute 'qualified_only'}
{attribute 'strict'}
TYPE E_RedPeer :		// 상대 PLC 상태 (EAP 하트비트 + 접점 신호로 판정. FB_RedPeerMonitor)
(
	Unknown		:= 0,	// 시작 직후: 아직 어느 쪽 신호도 못 봤고 시작 대기(tStartGrace) 안
	Alive		:= 1,	// EAP·접점 둘 다 살아 있음
	EapLost		:= 2,	// 접점만 살아 있음 = 통신(EAP) 고장. 상대는 살아 있음 (절체 조건 아님)
	WireLost	:= 3,	// EAP만 살아 있음 = 접점(배선) 고장. 상대는 살아 있음 (절체 조건 아님)
	Lost		:= 4	// 둘 다 끊김 = 상대 정지로 봄 (절체 조건)
) INT;
END_TYPE

// ---- 10_Core/90_Redundancy/ST_RedHeartbeat.TcDUT
TYPE ST_RedHeartbeat :		// 이중화 하트비트: 두 PLC가 EAP로 서로에게 매 스캔 보냄 (FB_RedLink). 필드를 바꾸면 두 PLC의 EAP 변수 연결도 같이 바꿈
STRUCT
	nProtoVer	: UINT := 2;	// 형식 번호. 상대와 다르면 필드 뜻이 다름
	nCounter	: UDINT;		// 보낼 때마다 1 증가. 상대가 이 값이 바뀌는지로 살아 있음을 봄
	nRole		: INT;			// 보낸 PLC의 역할 (E_RedRole)
	bActive		: BOOL;			// 보낸 PLC가 지금 장비에 쓰는가 (GVL_IF.g_bRedActive)
	nState		: INT;			// 보낸 PLC의 이중화 상태 (E_RedState). Primary가 Handover이면 Secondary가 Active를 내려놓음
END_STRUCT
END_TYPE

// ---- 10_Core/90_Redundancy/E_RedState.TcDUT
{attribute 'qualified_only'}
{attribute 'strict'}
TYPE E_RedState :		// 이 PLC의 이중화 상태 (FB_RedState). 역할(Primary/Secondary)은 고정 신분이고, 이 상태가 지금 장비에 쓰는지를 정함
(
	Init		:= 0,	// 시작 직후: 역할을 읽는 중이거나 상대 상태를 아직 모름. 장비에 쓰지 않음
	Standby		:= 1,	// 대기: 계산만 하고 장비에 쓰지 않음
	Active		:= 2,	// 장비에 씀 (GVL_IF.g_bRedActive = TRUE)
	Failed		:= 3,	// 설정 오류(Net ID 불일치·두 PLC 역할 같음). 장비에 쓰지 않음
	Handover	:= 4	// Primary 복귀 중: Secondary가 Active를 내려놓기를 기다림. 아직 장비에 쓰지 않음
) INT;
END_TYPE

// ---- 10_Core/90_Redundancy/E_RedSwitch.TcDUT
{attribute 'qualified_only'}
{attribute 'strict'}
TYPE E_RedSwitch :		// Active가 바뀐 마지막 이유 (FB_RedState)
(
	None		:= 0,	// 아직 없음
	Start		:= 1,	// 시작하면서 Active가 됨 (상대가 Active가 아님)
	PeerLost	:= 2,	// 절체: 상대가 Lost라 Secondary가 Active가 됨
	Failback	:= 3,	// 복귀: Primary가 Secondary에게서 Active를 넘겨받음
	Yield		:= 4	// 양보: Secondary가 Active를 내려놓음 (Primary가 돌아옴·동시 Active)
) INT;
END_TYPE

// ---- 10_Core/90_Redundancy/ST_RedSyncCfg.TcDUT
TYPE ST_RedSyncCfg :		// 동기화할 운영 설정 (GVL_PERSIST와 같은 모양. 모듈 설정 묶음 g_stModuleSet은 HMI가 두 PLC에 쓰므로 제외). 두 PLC가 EAP로 서로에게 매 스캔 보냄 (FB_RedSync). 필드를 바꾸면 두 PLC의 EAP 변수도 같이 바꿈
STRUCT
	nProtoVer		: UINT := 4;	// 형식 번호 (2: UPS 항목 추가 v2.43, 3: 사고 대응 된 동작 v2.49, 4: UPS 보관값 14칸·512 B 고정 v2.51. 두 PLC 프로그램이 달라 번호가 다르면 받은 값을 쓰지 않음)
	nSeq			: UDINT;		// 보낼 때마다 1 증가. 상대가 이 값이 바뀌는지로 살아 있음을 봄
	nModeReq1		: UINT;			// 제어 모드 요청 접속점 그룹 1 (GVL_SITE.g_fbCtrlMode1.i_nModeReq). [16번 수정 2026-11-09: nModeReq2(PCS2) 없앰]
	aeOpMode		: ARRAY[1..GVL_PARAM.UNIT_COUNT] OF E_OpMode;
	astGroupSet		: ARRAY[1..GVL_PARAM.GROUP_COUNT] OF ST_GroupSet;
	astManualPolicy	: ARRAY[1..GVL_PARAM.GROUP_COUNT] OF ST_ManualPolicy;
	astSourceReg	: ARRAY[1..GVL_PARAM.SOURCE_COUNT] OF ST_SourceReg;
	astLimitReg		: ARRAY[1..GVL_PARAM.LIMIT_COUNT] OF ST_ModuleReg;
	astPermitReg	: ARRAY[1..GVL_PARAM.PERMIT_COUNT] OF ST_ModuleReg;
	astCompReg		: ARRAY[1..GVL_PARAM.COMP_COUNT] OF ST_ModuleReg;
	astRuleCfg		: ARRAY[1..GVL_PARAM.RULE_COUNT] OF ST_RuleCfg;
	astOutputCfg	: ARRAY[1..GVL_PARAM.OUTPUT_COUNT] OF ST_OutputCfg;
	astUnitRuleReg	: ARRAY[1..GVL_PARAM.UNIT_RULE_COUNT] OF ST_RuleTargetReg;
	astBatRuleReg	: ARRAY[1..GVL_PARAM.BAT_RULE_COUNT] OF ST_RuleTargetReg;
	stCmdFilter		: ST_CmdFilterSet;
	stManualCmdSet	: ST_ManualCmdSet;
	stSeqSet		: ST_SeqSet;
	stBrokerWatch	: ST_BrokerWatchSet;	// MQTT 브로커 끊김 감시 [9번 수정 2026-11-09: 추가]
	astUpsDesired	: ARRAY[1..GVL_PARAM.UPS_COUNT] OF ST_UpsDesiredSet;	// UPS 설정 보관값 (GVL_PERSIST.g_astUpsDesired, 명세 RED-01 v2.43)
	bUpsSafetyRespEnable : BOOL;	// 사고·고장 대응 스위치 (GVL_PERSIST.g_bUpsSafetyRespEnable, 명세 RED-01 v2.43)
	awUpsRespDone	: ARRAY[1..GVL_PARAM.UPS_COUNT] OF WORD;	// 사고 대응 된 동작 비트 (FB_UpsSafetyResponse.q_wDone, GVL_IF.g_awUpsRespDone). 설정이 아님: 대기 쪽이 기억만 함 (명세 RED-01 v2.49)
	abSpare			: ARRAY[0..27] OF BYTE;	// 남는 자리: 전체를 512 B로 맞춤 (XAE EAP RedSyncCfg = ARRAY [0..511] OF BYTE). 위에 칸을 늘리면 이만큼 줄여 512 B 유지 (명세 RED-01 v2.51)
END_STRUCT
END_TYPE

// ---- 20_Module/Ups/E_UpsResult.TcDUT
// UPS·BMS 드라이버의 쓰기 요청 처리 결과.
{attribute 'qualified_only'}
{attribute 'strict'}
TYPE E_UpsResult : (
	None := 0, // 결과 없음
	Accepted := 1, // 요청 접수
	Disabled := 2, // 쓰기 비활성
	Busy := 3, // 다른 요청 처리 중
	Unsupported := 4, // 지원하지 않는 요청
	BadConfig := 5, // 설정값 오류
	WrongDevice := 6, // 대상 장치 불일치
	RevisionConflict := 7, // 설정 버전 불일치
	BadRequest := 8, // 잘못된 요청
	Duplicate := 9, // 중복 요청
	CommUnavailable := 10 // 통신 불가
) INT;
END_TYPE

// ---- 20_Module/Driver/Sebang/E_UpsCommand.TcDUT
// 세방 UPS 명령 주소. 해당 주소에 0x55를 쓰면 실행된다.
// BMS 명령 레지스터에 0x55를 쓰면 안 된다 (방식이 다름).
{attribute 'qualified_only'}
{attribute 'strict'}
TYPE E_UpsCommand : (
	Reset := 100, // 리셋
	BuzzerStop := 101, // 부저 정지
	RectifierOn := 102, // 정류기 ON
	RectifierOff := 103, // 정류기 OFF
	InverterOn := 104, // 인버터 ON
	InverterOff := 105, // 인버터 OFF
	BbcOn := 106, // BBC ON
	BbcOff := 107, // BBC OFF
	ToInverter := 108, // 인버터 절체
	ToBypass := 109, // 바이패스 절체 (BBC 대기 아님)
	FloatCharge := 110, // 부동충전
	EqualCharge := 111, // 균등충전
	AutoOn := 112, // 자동운전 ON
	AutoOff := 113, // 자동운전 OFF
	EmergencyDischarge := 114, // 비상 방전 시작
	PeriodicDischarge := 115, // 주기적 방전 시작
	PulseDischarge := 116, // 펄스 방전 시작
	CancelDischarge := 117, // 비상·주기적·펄스 방전 취소
	TrickleOn := 118, // 간헐충전 시작
	TrickleOff := 119, // 간헐충전 취소
	TemperatureOn := 120, // 온도보상 시작
	TemperatureOff := 121, // 온도보상 취소
	EcoOn := 122, // ECO ON
	EcoOff := 123, // ECO OFF
	PrltOn := 124, // PRLT ON
	PrltOff := 125 // PRLT OFF
) INT;
END_TYPE

// ---- 20_Module/Driver/Esolution/E_EsolutionOperation.TcDUT
{attribute 'qualified_only'}
{attribute 'strict'}
TYPE E_EsolutionOperation : (
	EmergencyStart := 0,
	PeriodicStart := 1,
	PulseStart := 2,
	DischargeCancel := 3,
	TrickleStart := 4,
	TrickleCancel := 5,
	TemperatureStart := 6,
	TemperatureCancel := 7,
	EcoStart := 8,
	EcoCancel := 9
) INT;
END_TYPE

// ---- 20_Module/Driver/Sebang/ST_UpsRaw.TcDUT
// 세방 UPS에서 읽은 변환 전 원본 값.
TYPE ST_UpsRaw :
STRUCT
	awInput : ARRAY[0..53] OF WORD; // FC04 Input 주소 0~53 (계측, 알람, 상태)
	awParam : ARRAY[0..66] OF WORD; // FC03 Holding 주소 0~66 (설정값)
END_STRUCT
END_TYPE

// ---- 20_Module/Ups/ST_UpsState.TcDUT
// UPS에서 읽어 공학 단위로 변환한 현재 상태.
// F_DecodeSebangUps가 ST_UpsRaw를 변환해 채우고, 알고리즘과 보고가 이 구조체를 읽는다.
TYPE ST_UpsState :
STRUCT

// UPS Metering Data 주소 순서
	fInputVoltageRV : REAL; // 0. 입력 선간 전압 R (V)
	fInputVoltageSV : REAL; // 1. 입력 선간 전압 S (V)
	fInputVoltageTV : REAL; // 2. 입력 선간 전압 T (V)
	fInputFrequencyHz : REAL; // 3. 입력 주파수 (Hz)
	fInputCurrentRA : REAL; // 4. 입력 전류 R (A)
	fInputCurrentSA : REAL; // 5. 입력 전류 S (A)
	fInputCurrentTA : REAL; // 6. 입력 전류 T (A)
	fInverterVoltageRV : REAL; // 7. 인버터 선간 전압 R (V)
	fInverterVoltageSV : REAL; // 8. 인버터 선간 전압 S (V)
	fInverterVoltageTV : REAL; // 9. 인버터 선간 전압 T (V)
	fInverterCurrentRA : REAL; // 10. 인버터 전류 R (A)
	fInverterCurrentSA : REAL; // 11. 인버터 전류 S (A)
	fInverterCurrentTA : REAL; // 12. 인버터 전류 T (A)
	fBypassVoltageRV : REAL; // 13. 바이패스 선간 전압 R (V)
	fBypassVoltageSV : REAL; // 14. 바이패스 선간 전압 S (V)
	fBypassVoltageTV : REAL; // 15. 바이패스 선간 전압 T (V)
	fBypassFrequencyHz : REAL; // 16. 바이패스 주파수 (Hz)
	fOutputVoltageRV : REAL; // 17. 출력 선간 전압 R (V)
	fOutputVoltageSV : REAL; // 18. 출력 선간 전압 S (V)
	fOutputVoltageTV : REAL; // 19. 출력 선간 전압 T (V)
	fOutputFrequencyHz : REAL; // 20. 출력 주파수 (Hz)
	fOutputCurrentRA : REAL; // 21. 출력 전류 R (A)
	fOutputCurrentSA : REAL; // 22. 출력 전류 S (A)
	fOutputCurrentTA : REAL; // 23. 출력 전류 T (A)
	fDcLinkVoltageV : REAL; // 24. DC 링크 전압 (V)
	fDcLinkHighVoltageV : REAL; // 25. DC 링크 상단 전압 (V)
	fDcLinkLowVoltageV : REAL; // 26. DC 링크 하단 전압 (V)
	fBatteryVoltageV : REAL; // 27. 배터리 전압 (V)
	fBatteryCurrentA : REAL; // 28. 배터리 전류 (A)
	fMpiCurrentAA : REAL; // 29. MPI A상 전류 (A)
	fMpiCurrentBA : REAL; // 30. MPI B상 전류 (A)
	fMpiCurrentCA : REAL; // 31. MPI C상 전류 (A)
	fInputApparentPowerKva : REAL; // 32. 입력 피상 전력 (kVA)
	fOutputApparentPowerKva : REAL; // 33. 출력 피상 전력 (kVA)
	fOutputActivePowerKw : REAL; // 34. 출력 유효 전력 (kW)
	// 주소 35~37: 예약 영역
	fTemperature1C : REAL; // 38. 온도 1 (℃)
	fTemperature2C : REAL; // 39. 온도 2 (℃)
	fTemperature3C : REAL; // 40. 온도 3 (℃)
	fTemperature4C : REAL; // 41. 온도 4 (℃)
	fTemperature5C : REAL; // 42. 온도 5 (℃)
	fBatteryRoomTemperatureC : REAL; // 43. 온도 6 / 배터리실 온도 (℃)
	wInputAlarm : WORD; // 44. 입력 알람
	wRectAlarm : WORD; // 45. 정류기 알람
	wBbcAlarm : WORD; // 46. 배터리 컨버터 알람
	wOutputAlarm : WORD; // 47. 출력 알람
	wInverterAlarm : WORD; // 48. 인버터 알람
	wBypassAlarm : WORD; // 49. 바이패스 알람
	wStatus1 : WORD; // 50. 상태 워드 1
	wStatus2 : WORD; // 51. 상태 워드 2
	fHmiVersion : REAL; // 52. HMI 버전
	fDspVersion : REAL; // 53. DSP 버전

// 해석한 운전 상태
	nBatMode : UINT; // 배터리 운전 모드
	bRectOn : BOOL; // 정류기 운전
	bRectNormal : BOOL; // 정류기 정상
	bBbcOn : BOOL; // 배터리 컨버터 운전
	bBbcNormal : BOOL; // 배터리 컨버터 정상
	bInverterOn : BOOL; // 인버터 운전
	bInverterNormal : BOOL; // 인버터 정상
	bOnBypass : BOOL; // 바이패스 공급
	bOnInverter : BOOL; // 인버터 공급
	bTemperatureEnabled : BOOL; // 온도보상 활성
	bBmsMinor : BOOL; // BMS 경고장
	bBmsMajor : BOOL; // BMS 중고장
	bEmergencyStop : BOOL; // 비상 정지
	awAlarmStatus : ARRAY[0..7] OF WORD; // 주소 44~51 알람·상태 묶음
	wOpCode : WORD; // H11 OP-CODE (설정값, Read Only). b3 Batt CB Trip = 배터리 MCCB Trip (명세 RD-UPS-01 v2.50)

// 프로그램 상태
	bComm : BOOL; // 통신 정상
	bValid : BOOL; // 데이터 유효
	bWriteFail : BOOL; // 쓰기 실패
	nSampleSeq : UDINT; // 표본 갱신 번호

END_STRUCT
END_TYPE

// ---- 20_Module/Driver/Esolution/ST_EsolutionRaw.TcDUT
TYPE ST_EsolutionRaw :
STRUCT

	awSystem : ARRAY[0..26] OF WORD; // Input 30001~30027 (맵 v1.4: 26 System Contactor State, 27 Rack Contactor State) [2026-11-13]
	awRackAnalog : ARRAY[0..39] OF WORD;
	awRackStatus : ARRAY[0..89] OF WORD;
	aawDetail : ARRAY[1..10,0..405] OF WORD;

END_STRUCT
END_TYPE

// ---- 20_Module/Driver/Esolution/ST_EsolutionState.TcDUT
TYPE ST_EsolutionState :
STRUCT

// System Data 1~25
	nHeartbeat : WORD; // 1. 하트비트
	fVoltageV : REAL; // 2. 전체 전압 (V)
	fCurrentA : REAL; // 3. 전체 전류 (A)
	fSocPct : REAL; // 4. 충전 상태 (%)
	fSohPct : REAL; // 5. 건강 상태 (%)
	fChargePowerKw : REAL; // 6. 충전 전력 (kW)
	fDischargePowerKw : REAL; // 7. 방전 전력 (kW)
	fMaxCellVoltageMv : REAL; // 8. 최대 셀 전압 (mV)
	fMinCellVoltageMv : REAL; // 9. 최소 셀 전압 (mV)
	fAvgCellVoltageMv : REAL; // 10. 평균 셀 전압 (mV)
	nMaxCellVoltageLocation : WORD; // 11. 최대 셀 전압 위치
	nMinCellVoltageLocation : WORD; // 12. 최소 셀 전압 위치
	fMaxCellTemperatureC : REAL; // 13. 최고 셀 온도 (℃)
	fMinCellTemperatureC : REAL; // 14. 최저 셀 온도 (℃)
	fAvgCellTemperatureC : REAL; // 15. 평균 셀 온도 (℃)
	nMaxCellTemperatureLocation : WORD; // 16. 최고 셀 온도 위치
	nMinCellTemperatureLocation : WORD; // 17. 최저 셀 온도 위치
	fMaxRackSocPct : REAL; // 18. 최대 랙 SOC (%)
	fMinRackSocPct : REAL; // 19. 최소 랙 SOC (%)
	fMaxRackVoltageV : REAL; // 20. 최대 랙 전압 (V)
	fMinRackVoltageV : REAL; // 21. 최소 랙 전압 (V)
	fChargeLimitKw : REAL; // 22. 충전 허용 전력 (kW)
	fDischargeLimitKw : REAL; // 23. 방전 허용 전력 (kW)
	fChargeCurrentLimitA : REAL; // 24. 충전 허용 전류 (A)
	fDischargeCurrentLimitA : REAL; // 25. 방전 허용 전류 (A)
// System Data 26~27 (맵 v1.4, 읽기 전용) [2026-11-13]
	wSystemContactor : WORD; // 26. 시스템 컨택터 상태 (b0 충전, b1 방전. 1 = 붙음)
	wRackContactor : WORD; // 27. 랙 컨택터 상태 (b0~b9 = 랙 1~10. 1 = 붙음)
	bChargeContactorClosed : BOOL; // 충전 컨택터 붙음 (26 b0)
	bDischargeContactorClosed : BOOL; // 방전 컨택터 붙음 (26 b1)

// 프로그램 상태
	bComm : BOOL; // 통신 정상
	bFresh : BOOL; // 데이터 갱신 정상
	bValid : BOOL; // 데이터 유효
	bWriteFail : BOOL; // 쓰기 실패
	bContactorFeedbackKnown : BOOL; // 컨택터 상태를 믿을 수 있음 (데이터 유효 = 맵 v1.4 26·27을 읽음)
	bWarn : BOOL; // 경보 발생
	bFault : BOOL; // 고장 발생
	bSystemLock : BOOL; // 시스템 잠금
	nSampleSeq : UDINT; // 표본 갱신 번호
	nRackCount : UINT; // 설치 랙 수
	nModuleCount : UINT; // 랙당 설치 모듈 수
	abDetailValid : ARRAY[1..10] OF BOOL; // 랙 상세 데이터 유효
	anDetailSeq : ARRAY[1..10] OF UDINT; // 랙 상세 갱신 번호

END_STRUCT
END_TYPE

// ---- 20_Module/Driver/Esolution/E_EsolutionControl.TcDUT
{attribute 'qualified_only'}
{attribute 'strict'}
TYPE E_EsolutionControl : (
	EmergencyShutdown := 11,
	SystemContactor := 12,	// 40013 Rack Contactor Control (맵 v1.4 이름): 1이면 랙 8개가 40001과 상관없이 한꺼번에 붙음
	ChargeContactor := 13,
	DischargeContactor := 14,
	ResetSystem := 30	// 40031 Reset System: 1이면 비상차단 해제 (명세 WR-BAT-01 v2.34)
) INT;
END_TYPE

// ---- 20_Module/Mqtt/Publish/ST_UpsPublish_V1.TcDUT
// UPS 1대의 MQTT 보고 데이터. 바이너리 구조라 필드 순서를 바꾸면 안 된다.
// 값은 FB_RptSebangUps가 ST_UpsState에서 복사한다.
{attribute 'pack_mode' := '1'}
TYPE ST_UpsPublish_V1 :
STRUCT
	DeviceIndex : UDINT; // UPS 번호 1~3
	SystemOperationMode : UDINT; // 시스템 운전모드 (enum) 0 수동, 1 모드스케줄. 출처 미정이라 지금은 0 [인터페이스 08.UPS 2026-11-12]
	OperationMode : UDINT; // 운전모드 (enum) 0 수동, 1 자동. EMS UPS 명령 101·102로 변경, 시작 기본값 1
	Status : UDINT; // b0 통신에러 b1 warning b2 fault b3 e-stop b4 충전 중(I50 b13 Batt charg Flag)
	UPS_ModeStatus : UDINT; // b0 부동충전 b1 균등충전 b2 대기 b3 주기적 방전 b4 펄스 방전 b5 간헐충전 (b0~b5 = I50 BAT Mode 값 0~5)
		// b6 비상 방전(I45 b8) b7 온도보상충전(I51 b2) b8 ECO(I48 b7) b9 PRLT(I50 b12) b10 Droop(I50 b11) b11 VSM(I45 b15) b12 Regen(I45 b8)
	MCCB_Status : UDINT; // b0 바이패스 M/C close b1 인버터 M/C close b2 입력 Pre M/C close b3 입력 M/C close b4 MBS C/B close b5 Out C/B Open b6 배터리 MCCB Trip (H11 b3, v2.50) (= I50 b1~b6, b5만 1이 개방)
	RectStatus : UDINT; // b0 정류부 기동(I45 b11) b1 정류부 정상(I45 b12) b2 Regen(I45 b8, 비상 방전)
	BBCStatus : UDINT; // b0 배터리 컨버터 기동(I46 b12) b1 배터리 컨버터 정상(I46 b13)
	InverterStatus : UDINT; // b0 인버터 기동(I48 b6) b1 인버터 정상(I48 b14) b2 인버터 출력(I48 b13 Load On Inverter)
	BypassStatus : UDINT; // b0 바이패스 출력(I48 b12 Load On Bypass)
	LineInputVoltage_R : REAL;
	LineInputVoltage_S : REAL;
	LineInputVoltage_T : REAL;
	InputFrequency : REAL;
	InputCurrent_R : REAL;
	InputCurrent_S : REAL;
	InputCurrent_T : REAL;
	InverterVoltage_R : REAL;
	InverterVoltage_S : REAL;
	InverterVoltage_T : REAL;
	InverterCurrent_R : REAL;
	InverterCurrent_S : REAL;
	InverterCurrent_T : REAL;
	BypassLineVoltage_R : REAL;
	BypassLineVoltage_S : REAL;
	BypassLineVoltage_T : REAL;
	BypassFrequency : REAL;
	LineOutputVoltage_R : REAL;
	LineOutputVoltage_S : REAL;
	LineOutputVoltage_T : REAL;
	FrequencyOutput : REAL;
	OutputCurrent_R : REAL;
	OutputCurrent_S : REAL;
	OutputCurrent_T : REAL;
	DcLinkVoltage : REAL;
	DcLinkVoltage_High : REAL;
	DcLinkVoltage_Low : REAL;
	BatteryVoltage : REAL;
	BatteryCurrent : REAL;
	MPI_A_Current : REAL;
	MPI_B_Current : REAL;
	MPI_C_Current : REAL;
	InputApparentPower : REAL;
	OutputApparentPower : REAL;
	OutputActivePower : REAL;
	Temp1 : REAL;
	Temp2 : REAL;
	Temp3 : REAL;
	Temp4 : REAL;
	Temp5 : REAL;
	Temp6 : REAL;
	// Warning·Fault: 회사 eventMap(001.UPS 경고장비트맵) 순서. 마스크로 거른 경고장·중고장을 맵 워드·비트 순서로 b0부터 빈칸 없이 (명세 RD-UPS-02 v2.20)
	Warning1 : UDINT; // 경고장 30개 b0~b29: I44 입력 → I45 정류부 → I46 BBC → I47 출력 → I49 바이패스 → I51 STATUS2
	Warning2 : UDINT; // 사용 안 함 (0)
	Warning3 : UDINT; // 사용 안 함 (0)
	Fault1 : UDINT; // 중고장 30개 b0~b29: I44 입력 → I45 정류부 → I46 BBC
	Fault2 : UDINT; // 중고장 19개 b0~b18: I47 출력 → I48 인버터 → I50 STATUS1 → I51 STATUS2
	Fault3 : UDINT; // 사용 안 함 (0)
END_STRUCT
END_TYPE

// ---- 20_Module/Mqtt/Publish/ST_ModulePublish_V1.TcDUT
{attribute 'pack_mode' := '1'}
TYPE ST_ModulePublish_V1 :
STRUCT
	BatIndex : UDINT;
	RackIndex : UDINT;
	DeviceIndex : UDINT;
	ModuleVolatge1 : REAL; // V. 인터페이스 10. Module.xlsx 표기 유지 (2026-11-17)
	ModuleVolatge2 : REAL; // V. BMS 맵에 별도 값 없음: 0
	ModuleVolatge3 : REAL; // V. BMS 맵에 별도 값 없음: 0
	ModuleTemp1 : REAL;
	ModuleTemp2 : REAL;
	ModuleTemp3 : REAL;
	CellVoltage1 : REAL;
	CellVoltage2 : REAL;
	CellVoltage3 : REAL;
	CellVoltage4 : REAL;
	CellVoltage5 : REAL;
	CellVoltage6 : REAL;
	CellVoltage7 : REAL;
	CellVoltage8 : REAL;
	CellVoltage9 : REAL;
	CellVoltage10 : REAL;
	CellVoltage11 : REAL;
	CellVoltage12 : REAL;
	CellVoltage13 : REAL;
	CellVoltage14 : REAL;
	CellVoltage15 : REAL;
	CellVoltage16 : REAL;
	CellVoltage17 : REAL;
	CellVoltage18 : REAL;
	CellVoltage19 : REAL;
	CellVoltage20 : REAL;
END_STRUCT
END_TYPE

// ---- 20_Module/Mqtt/Publish/ST_UpsPublishData.TcDUT
// EMS로 보내는 UPS MQTT 패킷 전체. 바이너리 구조라 필드 순서를 바꾸면 안 된다.
{attribute 'pack_mode' := '1'}
TYPE ST_UpsPublishData :
STRUCT
	Header : ST_MqttHeader; // MQTT 공통 헤더
	Devices : ARRAY[0..GVL_PARAM.UPS_COUNT-1] OF ST_UpsPublish_V1; // UPS별 데이터
END_STRUCT
END_TYPE

